    HMI_Message_Request : ARRAY[0..121] OF BOOL;  (* #HMI メッセージ表示要求; [0] 未使用; [1] 【Y616】A(左側) 供給スライド戻 異常表示; [2] 【Y617】A(左側) 供給スライド行 異常表示; [3] 【Y618】A(左側) 供給ピックアップ戻 異常表示; [4] 【Y619】A(左側) 供給ピックアップ行 異常表示; [5] 【Y620】A(左側) 供給チャック閉 戻 異常表示; [6] 【Y621】A(左側) 供給チャック開 行 異常表示; [7] 【Y622】B(右側) 供給スライド戻 異常表示; [8] 【Y623】B(右側) 供給スライド行 異常表示; [9] 【Y624】B(右側) 供給ピックアップ戻 異常表示; [10] 【Y625】B(右側) 供給ピックアップ行 異常表示; [11] 【Y626】B(右側) 供給チャック閉 戻 異常表示; [12] 【Y627】B(右側) 供給チャック開 行 異常表示; [13] 【Y700】A(左側) 高さ検査押え戻 異常表示; [14] 【Y701】A(左側) 高さ検査押え行 異常表示; [15] 【Y702】A(左側) 高さ検査持上戻 異常表示; [16] 【Y703】A(左側) 高さ検査持上行 異常表示; [17] 【Y704】A(左側) NG1ピックアップ戻 異常表示; [18] 【Y705】A(左側) NG1ピックアップ 行 異常表示; [19] 【Y706】A(左側) NG1チャック戻 異常表示; [20] 【Y707】A(左側) NG1チャック行 異常表示; [21] 【Y708】A(左側)ST4 反転1チャック閉 異常表示; [22] 【Y709】A(左側)ST4 反転1チャック開 異常表示; [23] 【Y710】A(左側)ST4 反転1ピックアップ戻 異常表示; [24] 【Y711】A(左側)ST4 反転1ピックアップ行 異常表示; [25] 【Y712】A(左側)ST6 反転2チャック閉 戻 異常表示; [26] 【Y713】A(左側)ST6 反転2チャック開 行 異常表示; [27] 【Y714】A(左側)ST6 反転2ピックアップ戻 異常表示; [28] 【Y715】A(左側)ST6 反転2ピックアップ行 異常表示; [29] 【Y716】A(左側) 排出チャック閉 戻 異常表示; [30] 【Y717】A(左側) 排出チャック開 行 異常表示; [31] 【Y718】A(左側) 排出フォルダ送り戻 異常表示; [32] 【Y719】A(左側) 排出フォルダ送り行 異常表示; [33] A(左側) 位置1ストッパー戻 異常表示; [34] 【Y720】A(左側) 位置1ストッパー 行 異常表示; [35] 【Y721】A(左側) 位置2ストッパー 異常表示; [36] 【Y721】A(左側) 位置2ストッパー 異常表示; [37] 【Y722】A(左側) 位置3ストッパー戻 異常表示; [38] 【Y722】A(左側) 位置3ストッパー行 異常表示; [39] Output_A_Error_M[33] 異常表示; [40] 【Y723】A(左側) 位置4ストッパー行 異常表示; [41] 【Y724】A(左側) 位置5ストッパー戻 異常表示; [42] 【Y724】A(左側) 位置5ストッパー行 異常表示; [43] 【Y725】A(左側) 位置6ストッパー戻 異常表示; [44] 【Y725】A(左側) 位置6ストッパー行 異常表示; [45] 【Y726】A(左側) ストックフォルダターン戻 異常表示; [46] 【Y727】A(左側) ストックフォルダターン行 異常表示; [47] 【Y728】A(左側) NG1仕分け 戻 異常表示; [48] 【Y729】A(左側) NG1仕分け 行 異常表示; [49] 【Y800】B(右側) 高さ検査押え戻 異常表示; [50] 【Y801】B(右側) 高さ検査押え行 異常表示; [51] 【Y802】B(右側) 高さ検査持上戻 異常表示; [52] 【Y803】B(右側) 高さ検査持上行 異常表示; [53] 【Y804】B(右側) NG1ピックアップ戻 異常表示; [54] 【Y805】B(右側) NG1ピックアップ 行 異常表示; [55] 【Y806】B(右側) NG1チャック戻 異常表示; [56] 【Y807】B(右側) NG1チャック行 異常表示; [57] 【Y808】B(右側)ST4 反転1チャック閉 戻 異常表示; [58] 【Y809】B(右側)ST4 反転1チャック開 戻 異常表示; [59] 【Y810】B(右側)ST4 反転1ピックアップ戻 異常表示; [60] 【Y811】B(右側)ST4 反転1ピックアップ行 異常表示; [61] 【Y812】B(右側)ST6 反転2チャック閉 戻 異常表示; [62] 【Y813】B(右側)ST6 反転2チャック開 行 異常表示; [63] 【Y814】B(右側)ST6 反転2ピックアップ戻 異常表示; [64] 【Y815】B(右側)ST6 反転2ピックアップ行 異常表示; [65] 【Y816】B(右側) 排出チャック閉 戻 異常表示; [66] 【Y817】B(右側) 排出チャック開 行 異常表示; [67] 【Y818】B(右側) 排出フォルダ送り戻 異常表示; [68] 【Y819】B(右側) 排出フォルダ送り行 異常表示; [69] 【Y820】B(右側) 位置1ストッパー 戻 異常表示; [70] 【Y820】B(右側) 位置1ストッパー 行 異常表示; [71] 【Y821】B(右側) 位置2ストッパー戻 異常表示; [72] 【Y821】B(右側) 位置2ストッパー行 異常表示; [73] 【Y822】B(右側) 位置3ストッパー戻 異常表示; [74] 【Y822】B(右側) 位置3ストッパー行 異常表示; [75] 【Y823】B(右側) 位置4ストッパー戻 異常表示; [76] 【Y823】B(右側) 位置4ストッパー行 異常表示; [77] 【Y824】B(右側) 位置5ストッパー戻 異常表示; [78] 【Y824】B(右側) 位置5ストッパー行 異常表示; [79] 【Y825】B(右側) 位置6ストッパー戻 異常表示; [80] 【Y825】B(右側) 位置6ストッパー行 異常表示; [81] 【Y826】B(右側) ストックフォルダターン戻 異常表示; [82] 【Y827】B(右側) ストックフォルダターン行 異常表示; [83] 【Y828】B(右側) NG1仕分け 戻 異常表示; [84] 【Y829】B(右側) NG1仕分け 行 異常表示; [85] 【Y1200】空コンテナ送り 戻 異常表示; [86] 【Y1201】空コンテナ送り 行 異常表示; [87] 【Y1202】段バラシ爪 戻 異常表示; [88] 【Y1203】段バラシ爪 行 異常表示; [89] 【Y1204】コンテナ排出 戻 異常表示; [90] 【Y1205】コンテナ排出 行 異常表示; [91] Output_Share_Error_M[7] 異常表示; [92] 【Y1207】箱入れチャック 行 異常表示; [93] 【Y1208】コンテナ仕分けストッパー 戻 異常表示; [94] 【Y1209】コンテナ仕分けストッパー 行 異常表示; [95] 【Y1210】コンテナ仕分け送り 戻 異常表示; [96] Output_Share_Error_M[12] 異常表示; [97] 【Y1300】A(左側) コンベア受渡送り戻 異常表示; [98] 【Y1301】A(左側) コンベア受渡送り行 異常表示; [99] 【Y1302】B(右側) コンベア受渡送り戻 異常表示; [100] 【Y1303】B(右側) コンベア受渡送り行 異常表示; [101] ST1 搬送ワーク不一致; [102] ST2 搬送ワーク不一致; [103] ST3 搬送ワーク不一致; [104] ST4 搬送ワーク不一致; [105] ST5 搬送ワーク不一致; [106] ST6 搬送ワーク不一致; [107] ST7 搬送ワーク不一致; [108] A(左側) ST1 FH測定時間超過; [109] A(左側) ST1 FH異常; [110] A(左側) ST5 FH異常; [111] B(右側) ST1 FH異常; [112] B(右側) ST5 FH異常; [113] A(左側) ST1 FH判定OK; [114] A(左側) ST1 FH判定NG1; [115] A(左側) ST1 FH判定NG2; [116] A(左側) ST1 検査前ワーク不一致; [117] A(左側) ST5 FH測定時間超過; [118] A(左側) ST5 FH判定OK; [119] A(左側) ST5 FH判定NG1; [120] A(左側) ST5 FH判定NG2; [121] A(左側) ST5 検査前ワーク不一致 *)
    HMI_Error_WorkSample : ARRAY[0..1] OF BOOL;  (* #HMI 再開前のワーク不一致; [0] A(左側) ST1; [1] A(左側) ST5 *)
    Error_ST1_A_Timeout : BOOL;  (* FHタイムアウト（非保持） *)
    Error_ST5_A_Timeout : BOOL;  (* FHタイムアウト（非保持） *)
    FH_B_ST1_Auto : BOOL;  (* B(右側) ST1 FH測定開始 *)
    Retry : ARRAY[0..99] OF BOOL;  (* 再試行：; [1] データ移動前 ワーク確; [4] ST3 検査前ワーク不一致エラー; [5] RCON1_1 機器異常; [6] A(左側) ST4 ワーク不一致エラー; [7] Stm A Axis000 絶対値位置決め エラー; [9] A(左側) ST6 ワーク不一致エラー; [10] Stm A Axis001 絶対値位置決め エラー; [12] RCON1_3 or 5機器異常 *)
    Stm_A_Rev_Axis000_MoveError : BOOL;  (* Stm A Axis000 絶対値位置決め エラー *)
    Stm_A_Rev1_Axis000_Power_Error : BOOL;  (* Stm A Axis000 サーボON エラー *)
    Stm_A_Rev_Axis001_MoveError : BOOL;  (* Stm A Axis001 絶対値位置決め エラー *)
    Stm_A_Rev2_Axis001_Power_Error : BOOL;  (* Stm A Axis001 サーボON エラー *)
    ST6_A_Rev2_End : BOOL;  (* ST6 A 動作完了 *)
    ST4_A_Rev_End : BOOL;  (* ST4 A 動作完了 *)
    RCON2_1_M : ARRAY[0..99] OF BOOL;  (* #RCON2_1 段バラシ; [1] 開始指令保持; [2] 予備 *)
    RCON2_1_IN_PositionDone : BOOL;  (* 位置決め完了 *)
    RCON2_1_IN_HomeDone : BOOL;  (* 原点復帰完了 *)
    RCON2_1_IN_Moving : BOOL;  (* 移動中 *)
    RCON2_1_IN_EmergencyStop : BOOL;  (* 非常停止状態（監視） *)
    RCON2_1_IN_ControllerReady : BOOL;  (* 準備完了 *)
    RCON2_1_IN_Zone2 : BOOL;  (* ゾーン2内 *)
    RCON2_1_IN_Zone1 : BOOL;  (* ゾーン1内 *)
    RCON2_1_IN_CommandDone : BOOL;  (* 指令完了 *)
    RCON2_1_IN_OverloadWarning : BOOL;  (* 過負荷警告 *)
    RCON2_1_IN_PushMiss : BOOL;  (* 押付け空振り（未使用） *)
    RCON2_1_IN_ServoReady : BOOL;  (* サーボON状態 *)
    RCON2_1_IN_Alarm : BOOL;  (* 軸異常 *)
    RCON2_1_Ready : BOOL;  (* 動作準備（安全許可とは別） *)
    RCON2_1_MoveDone : BOOL;  (* 動作完了 *)
    RCON2_1_OUT_TargetPos_mm : LREAL;  (* 目標位置 [mm] *)
    RCON2_1_OUT_PositionBand_mm : LREAL;  (* 位置決め幅 [mm] *)
    RCON2_1_OUT_Speed_mm_s : LREAL;  (* 指令速度 [mm/s] *)
    RCON2_1_OUT_AccDec_G : LREAL;  (* 加減速度 [G] *)
    RCON2_1_OUT_PushLimit_pct : LREAL;  (* 押付け制限 [%]（未使用） *)
    RCON2_1_ActualPos_mm : LREAL;  (* 現在位置 [mm] *)
    RCON2_1_Current_mA : DINT;  (* 指令電流 [mA]（監視値） *)
    RCON2_1_ActualSpeed_mm_s : LREAL;  (* 現在速度 [mm/s] *)
    RCON2_1_AlarmCode : UINT;  (* 軸異常コード *)
    RCON2_1_DataValid : BOOL;  (* 入力有効（安全許可とは別） *)
    RCON2_1_Auto : ARRAY[0..99] OF Bool;  (* 自動移動要求; [1] 初期動作① セイフティ; [2] 1段目 Pos; [3] 初期動作② セイフティ; [4] コンテナ排出 *)
    RCON2_2_M : ARRAY[0..99] OF BOOL;  (* #RCON2_2 箱詰めX; [1] 開始指令保持; [2] 今回移動受付：PEND OFF確認; [3] 自動開始許可 *)
    RCON2_2_IN_PositionDone : BOOL;  (* 位置決め完了 *)
    RCON2_2_IN_HomeDone : BOOL;  (* 原点復帰完了 *)
    RCON2_2_IN_Moving : BOOL;  (* 移動中 *)
    RCON2_2_IN_EmergencyStop : BOOL;  (* 非常停止状態（監視） *)
    RCON2_2_IN_ControllerReady : BOOL;  (* 準備完了 *)
    RCON2_2_IN_Zone2 : BOOL;  (* ゾーン2内 *)
    RCON2_2_IN_Zone1 : BOOL;  (* ゾーン1内 *)
    RCON2_2_IN_CommandDone : BOOL;  (* 指令完了 *)
    RCON2_2_IN_OverloadWarning : BOOL;  (* 過負荷警告 *)
    RCON2_2_IN_PushMiss : BOOL;  (* 押付け空振り（未使用） *)
    RCON2_2_IN_ServoReady : BOOL;  (* サーボON状態 *)
    RCON2_2_IN_Alarm : BOOL;  (* 軸異常 *)
    RCON2_2_Ready : BOOL;  (* 動作準備（安全許可とは別） *)
    RCON2_2_MoveDone : BOOL;  (* 動作完了 *)
    RCON2_2_OUT_TargetPos_mm : LREAL;  (* 目標位置 [mm] *)
    RCON2_2_OUT_PositionBand_mm : LREAL;  (* 位置決め幅 [mm] *)
    RCON2_2_OUT_Speed_mm_s : LREAL;  (* 指令速度 [mm/s] *)
    RCON2_2_OUT_AccDec_G : LREAL;  (* 加減速度 [G] *)
    RCON2_2_OUT_PushLimit_pct : LREAL;  (* 押付け制限 [%]（未使用） *)
    RCON2_2_ActualPos_mm : LREAL;  (* 現在位置 [mm] *)
    RCON2_2_Current_mA : DINT;  (* 指令電流 [mA]（監視値） *)
    RCON2_2_ActualSpeed_mm_s : LREAL;  (* 現在速度 [mm/s] *)
    RCON2_2_AlarmCode : UINT;  (* 軸異常コード *)
    RCON2_2_DataValid : BOOL;  (* 入力有効（安全許可とは別） *)
    RCON2_2_Auto : ARRAY[0..99] OF Bool;  (* 自動移動要求; [1] 自動要求1（未接続）; [2] 自動要求2（未接続）; [3] 自動要求3（未接続） *)
    RCON2_3_M : ARRAY[0..99] OF BOOL;  (* #RCON2_3 箱詰めY; [1] 開始指令保持; [2] 今回移動受付：PEND OFF確認; [3] 自動開始許可 *)
    RCON2_3_IN_PositionDone : BOOL;  (* 位置決め完了 *)
    RCON2_3_IN_HomeDone : BOOL;  (* 原点復帰完了 *)
    RCON2_3_IN_Moving : BOOL;  (* 移動中 *)
    RCON2_3_IN_EmergencyStop : BOOL;  (* 非常停止状態（監視） *)
    RCON2_3_IN_ControllerReady : BOOL;  (* 準備完了 *)
    RCON2_3_IN_Zone2 : BOOL;  (* ゾーン2内 *)
    RCON2_3_IN_Zone1 : BOOL;  (* ゾーン1内 *)
    RCON2_3_IN_CommandDone : BOOL;  (* 指令完了 *)
    RCON2_3_IN_OverloadWarning : BOOL;  (* 過負荷警告 *)
    RCON2_3_IN_PushMiss : BOOL;  (* 押付け空振り（未使用） *)
    RCON2_3_IN_ServoReady : BOOL;  (* サーボON状態 *)
    RCON2_3_IN_Alarm : BOOL;  (* 軸異常 *)
    RCON2_3_Ready : BOOL;  (* 動作準備（安全許可とは別） *)
    RCON2_3_MoveDone : BOOL;  (* 動作完了 *)
    RCON2_3_OUT_TargetPos_mm : LREAL;  (* 目標位置 [mm] *)
    RCON2_3_OUT_PositionBand_mm : LREAL;  (* 位置決め幅 [mm] *)
    RCON2_3_OUT_Speed_mm_s : LREAL;  (* 指令速度 [mm/s] *)
    RCON2_3_OUT_AccDec_G : LREAL;  (* 加減速度 [G] *)
    RCON2_3_OUT_PushLimit_pct : LREAL;  (* 押付け制限 [%]（未使用） *)
    RCON2_3_ActualPos_mm : LREAL;  (* 現在位置 [mm] *)
    RCON2_3_Current_mA : DINT;  (* 指令電流 [mA]（監視値） *)
    RCON2_3_ActualSpeed_mm_s : LREAL;  (* 現在速度 [mm/s] *)
    RCON2_3_AlarmCode : UINT;  (* 軸異常コード *)
    RCON2_3_DataValid : BOOL;  (* 入力有効（安全許可とは別） *)
    RCON2_3_Auto : ARRAY[0..99] OF Bool;  (* 自動移動要求; [1] 自動要求1（未接続）; [2] 自動要求2（未接続）; [3] 自動要求3（未接続） *)
    RCON2_4_M : ARRAY[0..99] OF BOOL;  (* #RCON2_4 箱詰めZ; [1] 開始指令保持; [2] 今回移動受付：PEND OFF確認; [3] 自動開始許可 *)
    RCON2_4_IN_PositionDone : BOOL;  (* 位置決め完了 *)
    RCON2_4_IN_HomeDone : BOOL;  (* 原点復帰完了 *)
    RCON2_4_IN_Moving : BOOL;  (* 移動中 *)
    RCON2_4_IN_EmergencyStop : BOOL;  (* 非常停止状態（監視） *)
    RCON2_4_IN_ControllerReady : BOOL;  (* 準備完了 *)
    RCON2_4_IN_Zone2 : BOOL;  (* ゾーン2内 *)
    RCON2_4_IN_Zone1 : BOOL;  (* ゾーン1内 *)
    RCON2_4_IN_CommandDone : BOOL;  (* 指令完了 *)
    RCON2_4_IN_OverloadWarning : BOOL;  (* 過負荷警告 *)
    RCON2_4_IN_PushMiss : BOOL;  (* 押付け空振り（未使用） *)
    RCON2_4_IN_ServoReady : BOOL;  (* サーボON状態 *)
    RCON2_4_IN_Alarm : BOOL;  (* 軸異常 *)
    RCON2_4_Ready : BOOL;  (* 動作準備（安全許可とは別） *)
    RCON2_4_MoveDone : BOOL;  (* 動作完了 *)
    RCON2_4_OUT_TargetPos_mm : LREAL;  (* 目標位置 [mm] *)
    RCON2_4_OUT_PositionBand_mm : LREAL;  (* 位置決め幅 [mm] *)
    RCON2_4_OUT_Speed_mm_s : LREAL;  (* 指令速度 [mm/s] *)
    RCON2_4_OUT_AccDec_G : LREAL;  (* 加減速度 [G] *)
    RCON2_4_OUT_PushLimit_pct : LREAL;  (* 押付け制限 [%]（未使用） *)
    RCON2_4_ActualPos_mm : LREAL;  (* 現在位置 [mm] *)
    RCON2_4_Current_mA : DINT;  (* 指令電流 [mA]（監視値） *)
    RCON2_4_ActualSpeed_mm_s : LREAL;  (* 現在速度 [mm/s] *)
    RCON2_4_AlarmCode : UINT;  (* 軸異常コード *)
    RCON2_4_DataValid : BOOL;  (* 入力有効（安全許可とは別） *)
    RCON2_4_Auto : ARRAY[0..99] OF Bool;  (* 自動移動要求; [1] 自動要求1（未接続）; [2] 自動要求2（未接続）; [3] 自動要求3（未接続） *)
    RCON2_5_M : ARRAY[0..99] OF BOOL;  (* #RCON2_5 コンテナ設置; [1] 開始指令保持; [2] 今回移動受付：PEND OFF確認; [3] 自動開始許可 *)
    RCON2_5_IN_PositionDone : BOOL;  (* 位置決め完了 *)
    RCON2_5_IN_HomeDone : BOOL;  (* 原点復帰完了 *)
    RCON2_5_IN_Moving : BOOL;  (* 移動中 *)
    RCON2_5_IN_EmergencyStop : BOOL;  (* 非常停止状態（監視） *)
    RCON2_5_IN_ControllerReady : BOOL;  (* 準備完了 *)
    RCON2_5_IN_Zone2 : BOOL;  (* ゾーン2内 *)
    RCON2_5_IN_Zone1 : BOOL;  (* ゾーン1内 *)
    RCON2_5_IN_CommandDone : BOOL;  (* 指令完了 *)
    RCON2_5_IN_OverloadWarning : BOOL;  (* 過負荷警告 *)
    RCON2_5_IN_PushMiss : BOOL;  (* 押付け空振り（未使用） *)
    RCON2_5_IN_ServoReady : BOOL;  (* サーボON状態 *)
    RCON2_5_IN_Alarm : BOOL;  (* 軸異常 *)
    RCON2_5_Ready : BOOL;  (* 動作準備（安全許可とは別） *)
    RCON2_5_MoveDone : BOOL;  (* 動作完了 *)
    RCON2_5_OUT_TargetPos_mm : LREAL;  (* 目標位置 [mm] *)
    RCON2_5_OUT_PositionBand_mm : LREAL;  (* 位置決め幅 [mm] *)
    RCON2_5_OUT_Speed_mm_s : LREAL;  (* 指令速度 [mm/s] *)
    RCON2_5_OUT_AccDec_G : LREAL;  (* 加減速度 [G] *)
    RCON2_5_OUT_PushLimit_pct : LREAL;  (* 押付け制限 [%]（未使用） *)
    RCON2_5_ActualPos_mm : LREAL;  (* 現在位置 [mm] *)
    RCON2_5_Current_mA : DINT;  (* 指令電流 [mA]（監視値） *)
    RCON2_5_ActualSpeed_mm_s : LREAL;  (* 現在速度 [mm/s] *)
    RCON2_5_AlarmCode : UINT;  (* 軸異常コード *)
    RCON2_5_DataValid : BOOL;  (* 入力有効（安全許可とは別） *)
    RCON2_5_Auto : ARRAY[0..99] OF Bool;  (* 自動移動要求; [1] コンテナトレイ方向NG; [2] 自動要求2（未接続）; [3] 自動要求3（未接続） *)
    Auto_Com_Start : BOOL;  (* 共通ユニット自動運転開始 *)
    Destacker_M : ARRAY[0..99] OF Bool;  (* 段バラシ工程; [5] 初回安全位置なし; [4] 初回安全位置あり; [2] 初回の爪保持; [3] 初回の位置判定; [6] 初回の爪戻し; [26] 初回確認済み; [27] 初回安全 前完了解除; [28] 初回1段 前完了解除; [29] 初回戻り 前完了解除; [30] 1段目 前完了解除; [31] 2段目 前完了解除; [32] 排出 前完了解除; [1] 初回確認開始; [7] 初回安全位置移動; [8] 初回1段目移動; [9] 初回コンテナ保持; [10] 初回安全位置戻り; [11] 初回の送り戻し; [12] 通常サイクル開始; [13] 送り戻り待ち; [14] コンテナ確認中; [15] コンテナ確認OK; [16] 1段目位置へ移動; [17] コンテナ切り離し; [18] 段積み判定; [19] 2段以上; [20] 1段のみ; [21] 2段目位置へ移動; [22] 上段コンテナ保持; [23] 安全・排出位置移動; [24] 送り行待ち; [25] 送り戻り待ち *)
    HMI_RCON2_1_OUT_TargetPos : ARRAY[0..99] OF LREAL;  (* 段バラシ 目標位置 [mm]; [1] ①④セイフティ・排出 Pos; [2] ②1段目 Pos; [3] ③2段目 Pos *)
    BoxPacking_Busy : BOOL;  (* 箱詰め動作中 *)
    Destacker_End : BOOL;  (* 1サイクル完了 *)
    Destacker_Error : BOOL;  (* 方向・1段目確認異常 *)
    Error_Destacker_M : ARRAY[0..99] OF Bool;  (* 段バラシエラー： *)
    ST7_B_SF_Wait_Pickup : BOOL;  (* フォルダストックB取出し待ち *)
END_VAR
VAR_GLOBAL RETAIN
    HMI_A_SF_StackPitch_mm : LREAL;  (* 左SF積みピッチ [mm] *)
END_VAR
VAR_GLOBAL
    A_Total_CT : INT;  (* A(左側)生産数 *)
    HMI_RCON2_4_OUT_TargetPos : ARRAY[0..99] OF LREAL;  (* 箱詰めZ：; [1] セイフティ 上昇 Pos; [2] フォルダストック 取出し降下Pos; [3] トレイ ワーク梱包 降下Pos *)
    Box_Total_CT : INT;  (* コンテナ入数 *)
END_VAR
VAR_GLOBAL RETAIN
    HMI_Box_X_Pitch_mm : LREAL;  (* 箱詰めX方向の1ピッチ [mm]：符号付き。正=座標増、負=座標減。使用前に設定。 *)
    HMI_Box_Y_Pitch_mm : LREAL;  (* 箱詰めY方向の1ピッチ [mm]：符号付き。正=座標増、負=座標減。使用前に設定。 *)
END_VAR

PROGRAM ModeManagement_モード管理
VAR
    Setting_M : BOOL;
    Manual_M : BOOL;
    Auto_M : BOOL;
    Dummy_M : BOOL;
    Inital_M : BOOL;
    Output_Error_M : ARRAY[0..99] OF Bool;
    Index_Error_001 : DINT;
    Index_B_001 : DINT;
    Index_Share_001 : DINT;
    Error_TON : ARRAY[0..99] OF TON;  (* [2] A(左側) ST1 測定タイムアウト; [4] A(左側) ST5 測定タイムアウト *)
    Error_TOF : ARRAY[0..99] OF TOF;
    AutoMode_A_M : ARRAY[0..99] OF Bool;
    ６ : DINT;
    ST4_A_Rev_01_Origin_M : ARRAY[0..99] OF Bool;  (* A(左側) ST4 反転1 原点復帰工程; [1] A(左側) ST4 反転1 原点復帰開始; [2] A(左側) ST4 反転1 原点復帰中; [3] A(左側) ST4 反転1 ピックアップ戻; [4] A(左側) ST4 反転1 モータ原点復帰開始; [5] A(左側) ST4 反転1 ピックアップ行; [6] A(左側) ST4 反転1 チャック閉; [7] A(左側) ST4 反転1 原点復帰完了（ワーク無） *)
    ST4_A_Rev_01_OriginDone : BOOL;  (* A(左側) ST4 反転1 原点復帰完了 *)
    ST4_A_Rev_02_Origin_M : ARRAY[0..99] OF Bool;  (* A(左側) ST6 反転2 原点復帰工程; [1] A(左側) ST6 反転2 原点復帰開始; [2] A(左側) ST6 反転2 原点復帰中; [3] A(左側) ST6 反転2 ピックアップ戻; [4] A(左側) ST6 反転2 モータ原点復帰開始; [5] A(左側) ST6 反転2 ピックアップ行; [6] A(左側) ST6 反転2 チャック閉; [7] A(左側) ST6 反転2 原点復帰完了（ワーク無） *)
    ST4_A_Rev_02_OriginDone : BOOL;  (* A(左側) ST6 反転2 原点復帰完了 *)
    ST4_B_Rev_01_Origin_M : ARRAY[0..99] OF Bool;  (* B(右側) ST4 反転1 原点復帰工程; [1] B(右側) ST4 反転1 原点復帰開始; [2] B(右側) ST4 反転1 原点復帰中; [3] B(右側) ST4 反転1 ピックアップ戻; [4] B(右側) ST4 反転1 モータ原点復帰開始; [5] B(右側) ST4 反転1 ピックアップ行; [6] B(右側) ST4 反転1 チャック閉; [7] B(右側) ST4 反転1 原点復帰完了（ワーク無） *)
    ST4_B_Rev_01_OriginDone : BOOL;  (* B(右側) ST4 反転1 原点復帰完了 *)
    ST4_B_Rev_02_Origin_M : ARRAY[0..99] OF Bool;  (* B(右側) ST6 反転2 原点復帰工程; [1] B(右側) ST6 反転2 原点復帰開始; [2] B(右側) ST6 反転2 原点復帰中; [3] B(右側) ST6 反転2 ピックアップ戻; [4] B(右側) ST6 反転2 モータ原点復帰開始; [5] B(右側) ST6 反転2 ピックアップ行; [6] B(右側) ST6 反転2 チャック閉; [7] B(右側) ST6 反転2 原点復帰完了（ワーク無） *)
    ST4_B_Rev_02_OriginDone : BOOL;  (* B(右側) ST6 反転2 原点復帰完了 *)
    ST1_B_Ca1_M : BOOL;
END_VAR
VAR_EXTERNAL
    Output_A_Error_M : ARRAY[0..99] OF Bool;
    Output_A_Restart_M : ARRAY[0..99] OF Bool;
    In_Sw_RESET : BOOL;
    In_Sw_START : BOOL;
    ManualMode : BOOL;
    M9999 : BOOL;
    Output_B_Error_M : ARRAY[0..99] OF Bool;  (* B(右側)シリンダエラー *)
    Output_B_Restart_M : ARRAY[0..99] OF Bool;  (* B(右側)シリンダ再開： *)
    Output_Share_Error_M : ARRAY[0..99] OF Bool;
    Output_Share_Restart_M : ARRAY[0..99] OF Bool;
    TimerQ_In_Sen_Accum_CV_A_Full : BOOL;
    Out_TDC_Stop : BOOL;
    In_Sen_Unl_Conv_A_Pass : BOOL;
    In_Sen_Accum_CV_A_Full : BOOL;
    In_Sen_Unl_Conv_B_Pass : BOOL;
    Pause : ARRAY[0..99] OF Bool;  (* [3] FH A(左側) ST1; [9] FH A(左側) ST5; [10] FH B(右側) ST1; [11] FH B(右側) ST5; [12] A(左側) ST6 反転2 ワーク不一致 *)
    AutoMode : BOOL;
    In_Sen_DOOR_01 : BOOL;
    In_Sen_DOOR_02 : BOOL;
    In_Sen_DOOR_03 : BOOL;
    In_Sen_DOOR_04 : BOOL;
    In_Sen_DOOR_05 : BOOL;
    In_Sen_DOOR_06 : BOOL;
    In_Sw_EMS1 : BOOL;
    In_Sw_EMS2 : BOOL;
    In_Sw_EMS3 : BOOL;
    In_Sen_AIR１_Pressure_01 : BOOL;
    In_Sen_AIR１_Pressure_02 : BOOL;
    In_Sen_AIR１_Pressure_03 : BOOL;
    TEST_M : ARRAY[0..99] OF Bool;
    ST0_Sup_Start : BOOL;  (* ST0_動作開始 *)
    Out_CYw_Sply_Pick_A_H_Auto : ARRAY[0..10] OF Bool;
    Out_CYw_Sply_Pick_A_H_Done : BOOL;
    Out_CYw_Sply_Slide_A_H_Auto : ARRAY[0..10] OF Bool;
    Out_CYw_Sply_Slide_A_H_Done : BOOL;
    Out_CYw_Sup_Chuck_A_Cl_H_Auto : ARRAY[0..10] OF Bool;
    Out_CYw_Sup_Chuck_A_Cl_H_Done : BOOL;
    In_Sen_Accum_CV_A_Arrival : BOOL;
    In_Sen_Work_A_Pos_00 : BOOL;
    Out_CYw_Sply_Pick_A_F_Auto : ARRAY[0..10] OF Bool;
    Out_CYw_Sply_Pick_A_F_Done : BOOL;
    Out_CYw_Sup_Chuck_A_Cl_F_Auto : ARRAY[0..10] OF Bool;
    Out_CYw_Sup_Chuck_A_Cl_F_Done : BOOL;
    Out_CYw_Sply_Slide_A_F_Auto : ARRAY[0..10] OF Bool;
    Out_CYw_Sply_Slide_A_F_Done : BOOL;
    Ins_A_Cv_Error : BOOL;
    Station_A_Data : ARRAY[0..8] OF sData;
    Ins_A_Cv_M : ARRAY[0..99] OF Bool;
    HMI_MessageNo : ARRAY[0..9] OF UINT;
    FH_A_ST1_Auto : BOOL;
    In_Sen_Accum_CV_B_Full : BOOL;
    FH_Line3_Error_Status_1 : BOOL;
    FH_Line0_Error_Status_1 : BOOL;
    FH_Line1_Error_Status_1 : BOOL;
    FH_Line2_Error_Status_1 : BOOL;
    FH_Line0_Error_Clear_1 : BOOL;
    FH_Line1_Error_Clear_1 : BOOL;
    FH_Line2_Error_Clear_1 : BOOL;
    FH_Line3_Error_Clear_1 : BOOL;
    Ins_A_Next_Cycle : BOOL;
    OriginDone : BOOL;  (* 原点復帰完了 *)
    DummyDone : BOOL;  (* ダミーチェック完了 *)
    HMI_CurrentPage : STRING[256];
    Ins_A_End : BOOL;
    Auto_A_Start : BOOL;  (* 自動運転 開始 *)
    Auto_Ready : BOOL;  (* 自動運転可能 *)
    ST0_A_Sup_Busy : BOOL;
    ST1_A_Ca1_Busy : BOOL;
    RCON1_1_IN_Alarm : BOOL;  (* 軸異常 *)
    RCON1_1_IN_EmergencyStop : BOOL;  (* 非常停止状態（監視） *)
    RCON1_1_Error : BOOL;  (* 異常予備（未接続） *)
    RCON1_1_IN_HomeDone : BOOL;  (* 原点復帰完了 *)
    RCON1_1_Error_Clear : BOOL;  (* 解除予備（未接続） *)
    Error_M : ARRAY[0..99] OF Bool;  (* エラー：; [1] シリンダ; [2] コンベア＆ドアセンサ; [3] 未使用：Error_ST1_A_M[0]へ移行; [4] A(左側)検査コンベア ワーク不一致; [5] 未使用：Error_ST3_A_M[1]へ移行; [9] 未使用：Error_ST5_A_M[0]へ移行; [10] 未使用：Error_ST1_B_M[0]へ移行; [11] 未使用：Error_ST5_B_M[0]へ移行; [12] 未使用：Error_ST6_A_M[0]へ移行 *)
    ST1_A_Ca1_M : ARRAY[0..99] OF Bool;  (* [6] A(左側) ST1 検査前ワーク不一致 *)
    ST2_A_Hgt_M : ARRAY[0..99] OF Bool;
    ST3_A_Dis1_M : ARRAY[0..99] OF Bool;
    HMI_Home_SW : BOOL;
    Origin_Busy : BOOL;  (* 原点復帰中 *)
    Out_CYw_Rev_01_Pick_A_H_Origin : ARRAY[0..10] OF Bool;  (* 原点復帰【Y710】A(左側)ST4 反転1ピックアップ戻： *)
    Out_CYw_Rev_01_Pick_A_H_Done : BOOL;  (* 【Y710】A(左側)ST4 反転1ピックアップ戻 動作完了 *)
    Stm_A_Rev_Axis000_Origin : BOOL;  (* A(左側) ST4 反転1 モータ原点復帰開始 *)
    Stm_A_Rev_Axis000_OriginDone : BOOL;  (* A(左側) ST4 反転1 モータ原点復帰完了 *)
    Out_CYw_Rev_01_Pick_A_F_Origin : ARRAY[0..99] OF Bool;  (* 原点復帰【Y711】A(左側)ST4 反転1ピックアップ行： *)
    Out_CYw_Rev_01_Pick_A_F_Done : BOOL;  (* 【Y711】A(左側)ST4 反転1ピックアップ行 動作完了 *)
    Out_CYw_Rev_01_Chk_A_H_Origin : ARRAY[0..99] OF Bool;  (* 原点復帰【Y708】A(左側)ST4 反転1チャック閉： *)
    Out_CYw_Rev_01_Chk_A_H_Done : BOOL;  (* 【Y708】A(左側)ST4 反転1チャック閉 動作完了 *)
    TimerQ_In_Sen_Work_A_Pos_04 : BOOL;
    Out_CYw_Rev_02_Pick_A_H_Origin : ARRAY[0..10] OF Bool;  (* 原点復帰 【Y714】A(左側)ST6 反転2ピックアップ戻 *)
    Out_CYw_Rev_02_Pick_A_H_Done : BOOL;  (* 【Y714】A(左側)ST6 反転2ピックアップ戻 動作完了 *)
    Stm_A_Rev_Axis001_Origin : BOOL;  (* A(左側) ST6 反転2 モータ原点復帰開始 *)
    Stm_A_Rev_Axis001_OriginDone : BOOL;  (* A(左側) ST6 反転2 モータ原点復帰完了 *)
    Out_CYw_Rev_02_Pick_A_F_Origin : ARRAY[0..99] OF Bool;  (* 原点復帰 【Y715】A(左側)ST6 反転2ピックアップ行 *)
    Out_CYw_Rev_02_Pick_A_F_Done : BOOL;  (* 【Y715】A(左側)ST6 反転2ピックアップ行 動作完了 *)
    Out_CYw_Rev_02_Chk_A_H_Origin : ARRAY[0..99] OF Bool;  (* 原点復帰 【Y712】A(左側)ST6 反転2チャック閉 戻 *)
    Out_CYw_Rev_02_Chk_A_H_Done : BOOL;  (* 【Y712】A(左側)ST6 反転2チャック閉 戻 動作完了 *)
    TimerQ_In_Sen_Work_A_Pos_06 : BOOL;  (* 【X208】A(左側)ワーク位置6 *)
    Auto_B_Start : BOOL;  (* B(右側)自動運転開始（後続処理未接続） *)
    Out_CYw_Rev_01_Pick_B_H_Origin : ARRAY[0..10] OF Bool;  (* 原点復帰 【Y810】B(右側)ST4 反転1ピックアップ戻 *)
    Out_CYw_Rev_01_Pick_B_H_Done : BOOL;  (* 【Y810】B(右側)ST4 反転1ピックアップ戻 動作完了 *)
    Stm_B_Rev_Axis002_Origin : BOOL;  (* B(右側) ST4 反転1 モータ原点復帰開始 *)
    Stm_B_Rev_Axis002_OriginDone : BOOL;  (* B(右側) ST4 反転1 モータ原点復帰完了 *)
    Out_CYw_Rev_01_Pick_B_F_Origin : ARRAY[0..99] OF Bool;  (* 原点復帰 【Y811】B(右側)ST4 反転1ピックアップ行 *)
    Out_CYw_Rev_01_Pick_B_F_Done : BOOL;  (* 【Y811】B(右側)ST4 反転1ピックアップ行 動作完了 *)
    Out_CYw_Rev_01_Chk_B_H_Origin : ARRAY[0..99] OF Bool;  (* 原点復帰 【Y808】B(右側)ST4 反転1チャック閉 戻 *)
    Out_CYw_Rev_01_Chk_B_H_Done : BOOL;  (* 【Y808】B(右側)ST4 反転1チャック閉 戻 動作完了 *)
    TimerQ_In_Sen_Work_B_Pos_04 : BOOL;  (* 【X406】B(右側)ワーク位置4 *)
    Out_CYw_Rev_02_Pick_B_H_Origin : ARRAY[0..10] OF Bool;  (* 原点復帰 【Y814】B(右側)ST6 反転2ピックアップ戻 *)
    Out_CYw_Rev_02_Pick_B_H_Done : BOOL;  (* 【Y814】B(右側)ST6 反転2ピックアップ戻 動作完了 *)
    Stm_B_Rev_Axis003_Origin : BOOL;  (* B(右側) ST6 反転2 モータ原点復帰開始 *)
    Stm_B_Rev_Axis003_OriginDone : BOOL;  (* B(右側) ST6 反転2 モータ原点復帰完了 *)
    Out_CYw_Rev_02_Pick_B_F_Origin : ARRAY[0..99] OF Bool;  (* 原点復帰 【Y815】B(右側)ST6 反転2ピックアップ行 *)
    Out_CYw_Rev_02_Pick_B_F_Done : BOOL;  (* 【Y815】B(右側)ST6 反転2ピックアップ行 動作完了 *)
    Out_CYw_Rev_02_Chk_B_H_Origin : ARRAY[0..99] OF Bool;  (* 原点復帰 【Y812】B(右側)ST6 反転2チャック閉 戻 *)
    Out_CYw_Rev_02_Chk_B_H_Done : BOOL;  (* 【Y812】B(右側)ST6 反転2チャック閉 戻 動作完了 *)
    TimerQ_In_Sen_Work_B_Pos_06 : BOOL;  (* 【X408】B(右側)ワーク位置6 *)
    ST4_A_Rev1_M : ARRAY[0..99] OF Bool;  (* [10] A(左側) ST4 ワーク不一致エラー; [12] 【Y708】A(左側) ST4 反転1チャック閉 *)
    ST5_A_Ca2_M : ARRAY[0..99] OF Bool;  (* A(左側) ST5 カメラ2工程; [1] A(左側) ST5 カメラ2検査開始; [2] 【Y724】A(左側) ST5 ストッパー戻; [3] A(左側) ST5 ワーク有無判定; [4] A(左側) ST5 ワーク有; [5] A(左側) ST5 ワーク無; [6] A(左側) ST5 検査前ワーク不一致; [7] A(左側) ST5 FH測定開始 *)
    FH_A_ST5_Auto : BOOL;  (* A(左側) ST5 FH自動測定 *)
END_VAR
VAR_EXTERNAL CONSTANT
    ST6_A_Rev2_M : ARRAY[0..99] OF Bool;  (* A(左側) ST6 反転2工程; [1] A(左側) ST6 反転2 動作開始; [2] A(左側) ST6 反転2 【Y714】ピックアップ戻; [3] A(左側) ST6 反転2 【Y725】位置6ストッパー戻; [4] A(左側) ST6 反転2 原点角度転送; [5] A(左側) ST6 反転2 原点位置移動開始; [6] A(左側) ST6 反転2 原点位置移動完了; [7] A(左側) ST6 反転2 ワーク有無判定; [8] A(左側) ST6 反転2 ワーク有・前工程OK; [9] A(左側) ST6 反転2 ワーク無・前工程NG; [10] A(左側) ST6 反転2 ワーク不一致エラー; [11] A(左側) ST6 反転2 【Y715】反転前ピックアップ行; [12] A(左側) ST6 反転2 【Y712】チャック閉; [13] A(左側) ST6 反転2 【Y714】反転前ピックアップ戻; [14] A(左側) ST6 反転2 反転角度転送; [15] A(左側) ST6 反転2 反転位置移動完了; [16] A(左側) ST6 反転2 【Y715】設置ピックアップ行; [17] A(左側) ST6 反転2 【Y713】チャック開; [18] A(左側) ST6 反転2 【Y714】設置ピックアップ戻 *)
END_VAR
VAR_EXTERNAL
    ST7_A_Dis2_M : ARRAY[0..99] OF Bool;  (* [9] ワーク有; [10] ワーク無; [11] 有無・NG満杯異常; [12] 回収下降位置転送; [13] 回収下降要求; [14] ワーク保持; [15] 保持後上昇位置転送; [16] 保持後上昇要求; [17] 仕分け位置選択; [18] OK選択; [19] キズNG選択; [20] 姿NG選択; [21] OK送り行開始; [22] 仕分け左右移動中; [23] 下降位置選択; [24] OK積み位置; [25] キズNG下降位置; [26] 姿NG下降位置; [27] 配置下降要求; [28] ワーク解放; [29] 解放後上昇位置転送; [30] 解放後上昇要求; [31] 左右原点位置転送; [32] 左右原点移動要求; [33] 最後の送り戻; [1] 排出動作開始; [2] 初期チャック戻; [3] 初期上昇位置転送; [4] 初期上昇要求; [5] 初期左右位置転送; [6] 初期左右移動要求; [7] 初期送り戻; [8] ワーク有無判定; [42] 今回ワーク加算済み; [43] 積み設定・判定異常; [44] フォルダ回転異常; [45] ワーク回収開始許可; [46] 今回の初期位置確認済み; [34] 初期上昇 前完了解除; [35] 初期左右 前完了解除; [36] 回収下降 前完了解除; [37] 保持後上昇 前完了解除; [38] 仕分け左右 前完了解除; [39] 配置下降 前完了解除; [40] 解放後上昇 前完了解除; [41] 左右戻り 前完了解除 *)
    Error_ST1_A_M : ARRAY[0..4] OF BOOL;  (* #A(左側) ST1 カメラ1 異常; [0] 総合異常; [1] 機器異常; [2] タイムアウト; [3] ワーク不一致; [4] 予備（監視なし） *)
    Error_ST1_B_M : ARRAY[0..4] OF BOOL;  (* #B(右側) ST1 カメラ1 異常; [0] 総合異常; [1] 機器異常; [2] 予備（監視なし）; [3] 予備（監視なし）; [4] 予備（監視なし） *)
    Error_ST2_A_M : ARRAY[0..4] OF BOOL;  (* #A(左側) ST2 高さ検査 異常; [0] 総合異常; [1] 予備（監視なし）; [2] 予備（監視なし）; [3] ワーク不一致; [4] 予備（監視なし） *)
    Error_ST3_A_M : ARRAY[0..4] OF BOOL;  (* #A(左側) ST3 NG1排出 異常; [0] 総合異常; [1] 機器異常; [2] 予備（監視なし）; [3] ワーク不一致; [4] 予備（監視なし） *)
    Error_ST4_A_M : ARRAY[0..4] OF BOOL;  (* #A(左側) ST4 反転1 異常; [0] 総合異常; [1] 予備（監視なし）; [2] 予備（監視なし）; [3] ワーク不一致; [4] 予備（監視なし） *)
    Error_ST5_A_M : ARRAY[0..4] OF BOOL;  (* #A(左側) ST5 カメラ2 異常; [0] 総合異常; [1] 機器異常; [2] タイムアウト; [3] ワーク不一致; [4] 予備（監視なし） *)
    Error_ST5_B_M : ARRAY[0..4] OF BOOL;  (* #B(右側) ST5 カメラ2 異常; [0] 総合異常; [1] 機器異常; [2] 予備（監視なし）; [3] 予備（監視なし）; [4] 予備（監視なし） *)
    Error_ST6_A_M : ARRAY[0..4] OF BOOL;  (* #A(左側) ST6 反転2 異常; [0] 総合異常; [1] 予備（監視なし）; [2] 予備（監視なし）; [3] ワーク不一致; [4] 予備（監視なし） *)
    Error_ST7_A_M : ARRAY[0..4] OF BOOL;  (* #A(左側) ST7 SF排出 異常; [0] 総合異常; [1] 予備（監視なし）; [2] 予備（監視なし）; [3] ワーク不一致; [4] 満杯 *)
    Error_ST7_A_Source_M : ARRAY[0..4] OF BOOL;  (* #A(左側) ST7 発生理由（内部保持）; [3] ワーク不一致; [4] 満杯（既存B側入力） *)
    HMI_Message_Request : ARRAY[0..121] OF BOOL;  (* #HMI メッセージ表示要求; [0] 未使用; [1] 【Y616】A(左側) 供給スライド戻 異常表示; [2] 【Y617】A(左側) 供給スライド行 異常表示; [3] 【Y618】A(左側) 供給ピックアップ戻 異常表示; [4] 【Y619】A(左側) 供給ピックアップ行 異常表示; [5] 【Y620】A(左側) 供給チャック閉 戻 異常表示; [6] 【Y621】A(左側) 供給チャック開 行 異常表示; [7] 【Y622】B(右側) 供給スライド戻 異常表示; [8] 【Y623】B(右側) 供給スライド行 異常表示; [9] 【Y624】B(右側) 供給ピックアップ戻 異常表示; [10] 【Y625】B(右側) 供給ピックアップ行 異常表示; [11] 【Y626】B(右側) 供給チャック閉 戻 異常表示; [12] 【Y627】B(右側) 供給チャック開 行 異常表示; [13] 【Y700】A(左側) 高さ検査押え戻 異常表示; [14] 【Y701】A(左側) 高さ検査押え行 異常表示; [15] 【Y702】A(左側) 高さ検査持上戻 異常表示; [16] 【Y703】A(左側) 高さ検査持上行 異常表示; [17] 【Y704】A(左側) NG1ピックアップ戻 異常表示; [18] 【Y705】A(左側) NG1ピックアップ 行 異常表示; [19] 【Y706】A(左側) NG1チャック戻 異常表示; [20] 【Y707】A(左側) NG1チャック行 異常表示; [21] 【Y708】A(左側)ST4 反転1チャック閉 異常表示; [22] 【Y709】A(左側)ST4 反転1チャック開 異常表示; [23] 【Y710】A(左側)ST4 反転1ピックアップ戻 異常表示; [24] 【Y711】A(左側)ST4 反転1ピックアップ行 異常表示; [25] 【Y712】A(左側)ST6 反転2チャック閉 戻 異常表示; [26] 【Y713】A(左側)ST6 反転2チャック開 行 異常表示; [27] 【Y714】A(左側)ST6 反転2ピックアップ戻 異常表示; [28] 【Y715】A(左側)ST6 反転2ピックアップ行 異常表示; [29] 【Y716】A(左側) 排出チャック閉 戻 異常表示; [30] 【Y717】A(左側) 排出チャック開 行 異常表示; [31] 【Y718】A(左側) 排出フォルダ送り戻 異常表示; [32] 【Y719】A(左側) 排出フォルダ送り行 異常表示; [33] A(左側) 位置1ストッパー戻 異常表示; [34] 【Y720】A(左側) 位置1ストッパー 行 異常表示; [35] 【Y721】A(左側) 位置2ストッパー 異常表示; [36] 【Y721】A(左側) 位置2ストッパー 異常表示; [37] 【Y722】A(左側) 位置3ストッパー戻 異常表示; [38] 【Y722】A(左側) 位置3ストッパー行 異常表示; [39] Output_A_Error_M[33] 異常表示; [40] 【Y723】A(左側) 位置4ストッパー行 異常表示; [41] 【Y724】A(左側) 位置5ストッパー戻 異常表示; [42] 【Y724】A(左側) 位置5ストッパー行 異常表示; [43] 【Y725】A(左側) 位置6ストッパー戻 異常表示; [44] 【Y725】A(左側) 位置6ストッパー行 異常表示; [45] 【Y726】A(左側) ストックフォルダターン戻 異常表示; [46] 【Y727】A(左側) ストックフォルダターン行 異常表示; [47] 【Y728】A(左側) NG1仕分け 戻 異常表示; [48] 【Y729】A(左側) NG1仕分け 行 異常表示; [49] 【Y800】B(右側) 高さ検査押え戻 異常表示; [50] 【Y801】B(右側) 高さ検査押え行 異常表示; [51] 【Y802】B(右側) 高さ検査持上戻 異常表示; [52] 【Y803】B(右側) 高さ検査持上行 異常表示; [53] 【Y804】B(右側) NG1ピックアップ戻 異常表示; [54] 【Y805】B(右側) NG1ピックアップ 行 異常表示; [55] 【Y806】B(右側) NG1チャック戻 異常表示; [56] 【Y807】B(右側) NG1チャック行 異常表示; [57] 【Y808】B(右側)ST4 反転1チャック閉 戻 異常表示; [58] 【Y809】B(右側)ST4 反転1チャック開 戻 異常表示; [59] 【Y810】B(右側)ST4 反転1ピックアップ戻 異常表示; [60] 【Y811】B(右側)ST4 反転1ピックアップ行 異常表示; [61] 【Y812】B(右側)ST6 反転2チャック閉 戻 異常表示; [62] 【Y813】B(右側)ST6 反転2チャック開 行 異常表示; [63] 【Y814】B(右側)ST6 反転2ピックアップ戻 異常表示; [64] 【Y815】B(右側)ST6 反転2ピックアップ行 異常表示; [65] 【Y816】B(右側) 排出チャック閉 戻 異常表示; [66] 【Y817】B(右側) 排出チャック開 行 異常表示; [67] 【Y818】B(右側) 排出フォルダ送り戻 異常表示; [68] 【Y819】B(右側) 排出フォルダ送り行 異常表示; [69] 【Y820】B(右側) 位置1ストッパー 戻 異常表示; [70] 【Y820】B(右側) 位置1ストッパー 行 異常表示; [71] 【Y821】B(右側) 位置2ストッパー戻 異常表示; [72] 【Y821】B(右側) 位置2ストッパー行 異常表示; [73] 【Y822】B(右側) 位置3ストッパー戻 異常表示; [74] 【Y822】B(右側) 位置3ストッパー行 異常表示; [75] 【Y823】B(右側) 位置4ストッパー戻 異常表示; [76] 【Y823】B(右側) 位置4ストッパー行 異常表示; [77] 【Y824】B(右側) 位置5ストッパー戻 異常表示; [78] 【Y824】B(右側) 位置5ストッパー行 異常表示; [79] 【Y825】B(右側) 位置6ストッパー戻 異常表示; [80] 【Y825】B(右側) 位置6ストッパー行 異常表示; [81] 【Y826】B(右側) ストックフォルダターン戻 異常表示; [82] 【Y827】B(右側) ストックフォルダターン行 異常表示; [83] 【Y828】B(右側) NG1仕分け 戻 異常表示; [84] 【Y829】B(右側) NG1仕分け 行 異常表示; [85] 【Y1200】空コンテナ送り 戻 異常表示; [86] 【Y1201】空コンテナ送り 行 異常表示; [87] 【Y1202】段バラシ爪 戻 異常表示; [88] 【Y1203】段バラシ爪 行 異常表示; [89] 【Y1204】コンテナ排出 戻 異常表示; [90] 【Y1205】コンテナ排出 行 異常表示; [91] Output_Share_Error_M[7] 異常表示; [92] 【Y1207】箱入れチャック 行 異常表示; [93] 【Y1208】コンテナ仕分けストッパー 戻 異常表示; [94] 【Y1209】コンテナ仕分けストッパー 行 異常表示; [95] 【Y1210】コンテナ仕分け送り 戻 異常表示; [96] Output_Share_Error_M[12] 異常表示; [97] 【Y1300】A(左側) コンベア受渡送り戻 異常表示; [98] 【Y1301】A(左側) コンベア受渡送り行 異常表示; [99] 【Y1302】B(右側) コンベア受渡送り戻 異常表示; [100] 【Y1303】B(右側) コンベア受渡送り行 異常表示; [101] ST1 搬送ワーク不一致; [102] ST2 搬送ワーク不一致; [103] ST3 搬送ワーク不一致; [104] ST4 搬送ワーク不一致; [105] ST5 搬送ワーク不一致; [106] ST6 搬送ワーク不一致; [107] ST7 搬送ワーク不一致; [108] A(左側) ST1 FH測定時間超過; [109] A(左側) ST1 FH異常; [110] A(左側) ST5 FH異常; [111] B(右側) ST1 FH異常; [112] B(右側) ST5 FH異常; [113] A(左側) ST1 FH判定OK; [114] A(左側) ST1 FH判定NG1; [115] A(左側) ST1 FH判定NG2; [116] A(左側) ST1 検査前ワーク不一致; [117] A(左側) ST5 FH測定時間超過; [118] A(左側) ST5 FH判定OK; [119] A(左側) ST5 FH判定NG1; [120] A(左側) ST5 FH判定NG2; [121] A(左側) ST5 検査前ワーク不一致 *)
    HMI_Error_WorkSample : ARRAY[0..1] OF BOOL;  (* #HMI 再開前のワーク不一致; [0] A(左側) ST1; [1] A(左側) ST5 *)
    Error_ST1_A_Timeout : BOOL;  (* FHタイムアウト（非保持） *)
    Error_ST5_A_Timeout : BOOL;  (* FHタイムアウト（非保持） *)
    TimerQ_In_Sen_Work_A_Pos_07 : BOOL;  (* 【X209】A(左側)ワーク位置7 *)
    TimerQ_In_Sen_NG2_Tray_B_Full : BOOL;  (* 【X412】B(右側) NG2トレイ満杯停止 *)
    Retry : ARRAY[0..99] OF BOOL;
    Stm_A_Rev1_Axis000_Power_Error : BOOL;
    Stm_A_Rev_Axis000_MoveError : BOOL;
    RCON1_3_Error : BOOL;
    RCON1_3_Error_Clear : BOOL;
    RCON1_3_IN_Alarm : BOOL;
    RCON1_3_IN_EmergencyStop : BOOL;
    TimerQ_In_Sen_NG2_Tray_A_Full : BOOL;
    RCON1_5_Error : BOOL;
    RCON1_5_Error_Clear : BOOL;
    Auto_Com_Start : BOOL;  (* 共通ユニット自動運転開始 *)
    Destacker_Error : BOOL;  (* 方向・1段目確認異常 *)
    Error_Destacker_M : ARRAY[0..99] OF Bool;  (* 段バラシエラー： *)
END_VAR
VAR
    _p1 : BOOL;
    _p2 : BOOL;
    _p3 : BOOL;
    _p4 : BOOL;
    _p5 : BOOL;
    _p6 : BOOL;
    _p7 : BOOL;
    _p8 : BOOL;
    _p9 : BOOL;
    _p10 : BOOL;
    _p11 : BOOL;
    _p12 : BOOL;
    _p13 : BOOL;
    _p14 : BOOL;
    _p15 : BOOL;
    _p16 : BOOL;
    _p17 : BOOL;
    _p18 : BOOL;
    _p19 : BOOL;
    _p20 : BOOL;
    _p21 : BOOL;
    _p22 : BOOL;
    _p23 : BOOL;
    _p24 : BOOL;
    _e25 : R_TRIG;
    _e26 : R_TRIG;
    _e27 : R_TRIG;
    _e28 : R_TRIG;
    _e29 : R_TRIG;
    _e30 : R_TRIG;
    _e31 : R_TRIG;
    _e32 : R_TRIG;
    _e33 : R_TRIG;
    _e34 : R_TRIG;
    _p35 : BOOL;
    _p36 : BOOL;
    _p37 : BOOL;
    _e38 : R_TRIG;
    _e39 : R_TRIG;
    _e40 : R_TRIG;
    _e41 : R_TRIG;
    _e42 : R_TRIG;
    _e43 : R_TRIG;
    _e44 : R_TRIG;
    _e45 : R_TRIG;
    _e46 : R_TRIG;
    _e47 : R_TRIG;
    _p48 : BOOL;
END_VAR

(* Section Initial_初期化処理: ladder, written here as Structured Text *)

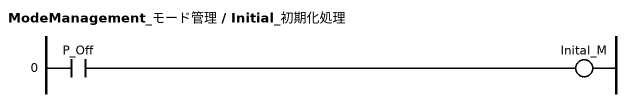
(* Rung 0 *)
Inital_M := P_Off;

(* Section Origin_原点復帰: ladder, written here as Structured Text *)

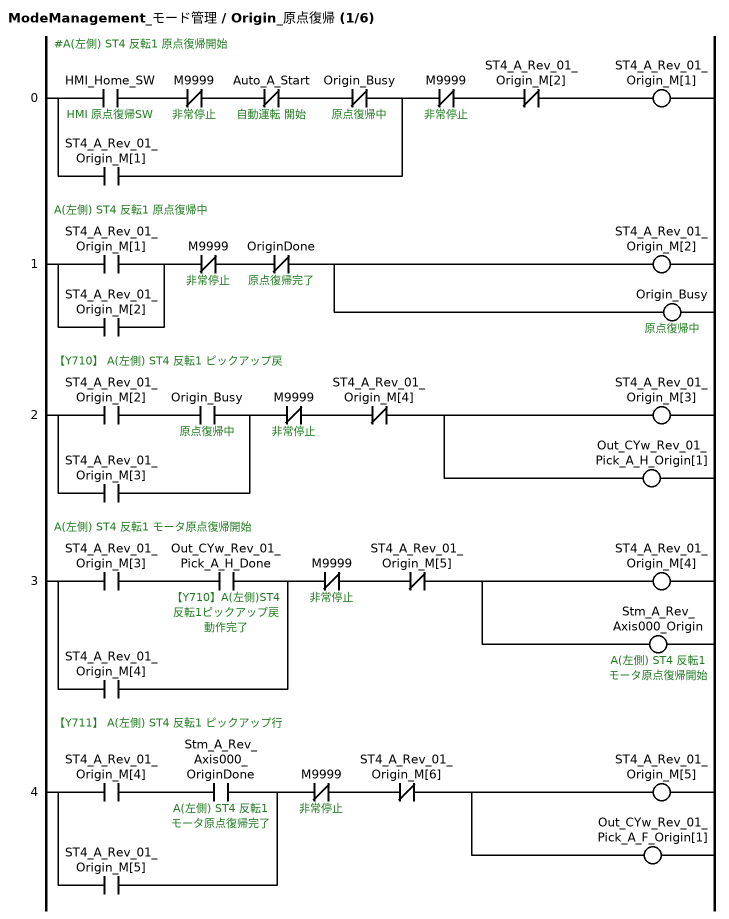
(* Rung 0: #A(左側) ST4 反転1 原点復帰開始 *)
ST4_A_Rev_01_Origin_M[1] := ((HMI_Home_SW AND NOT M9999 AND NOT Auto_A_Start AND NOT Origin_Busy) OR ST4_A_Rev_01_Origin_M[1]) AND NOT M9999 AND NOT ST4_A_Rev_01_Origin_M[2];
(* Rung 1: A(左側) ST4 反転1 原点復帰中 *)
_p1 := (ST4_A_Rev_01_Origin_M[1] OR ST4_A_Rev_01_Origin_M[2]) AND NOT M9999 AND NOT OriginDone;
ST4_A_Rev_01_Origin_M[2] := _p1;
Origin_Busy := _p1;
(* Rung 2: 【Y710】 A(左側) ST4 反転1 ピックアップ戻 *)
_p2 := ((ST4_A_Rev_01_Origin_M[2] AND Origin_Busy) OR ST4_A_Rev_01_Origin_M[3]) AND NOT M9999 AND NOT ST4_A_Rev_01_Origin_M[4];
ST4_A_Rev_01_Origin_M[3] := _p2;
Out_CYw_Rev_01_Pick_A_H_Origin[1] := _p2;
(* Rung 3: A(左側) ST4 反転1 モータ原点復帰開始 *)
_p3 := ((ST4_A_Rev_01_Origin_M[3] AND Out_CYw_Rev_01_Pick_A_H_Done) OR ST4_A_Rev_01_Origin_M[4]) AND NOT M9999 AND NOT ST4_A_Rev_01_Origin_M[5];
ST4_A_Rev_01_Origin_M[4] := _p3;
Stm_A_Rev_Axis000_Origin := _p3;
(* Rung 4: 【Y711】 A(左側) ST4 反転1 ピックアップ行 *)
_p4 := ((ST4_A_Rev_01_Origin_M[4] AND Stm_A_Rev_Axis000_OriginDone) OR ST4_A_Rev_01_Origin_M[5]) AND NOT M9999 AND NOT ST4_A_Rev_01_Origin_M[6];
ST4_A_Rev_01_Origin_M[5] := _p4;
Out_CYw_Rev_01_Pick_A_F_Origin[1] := _p4;

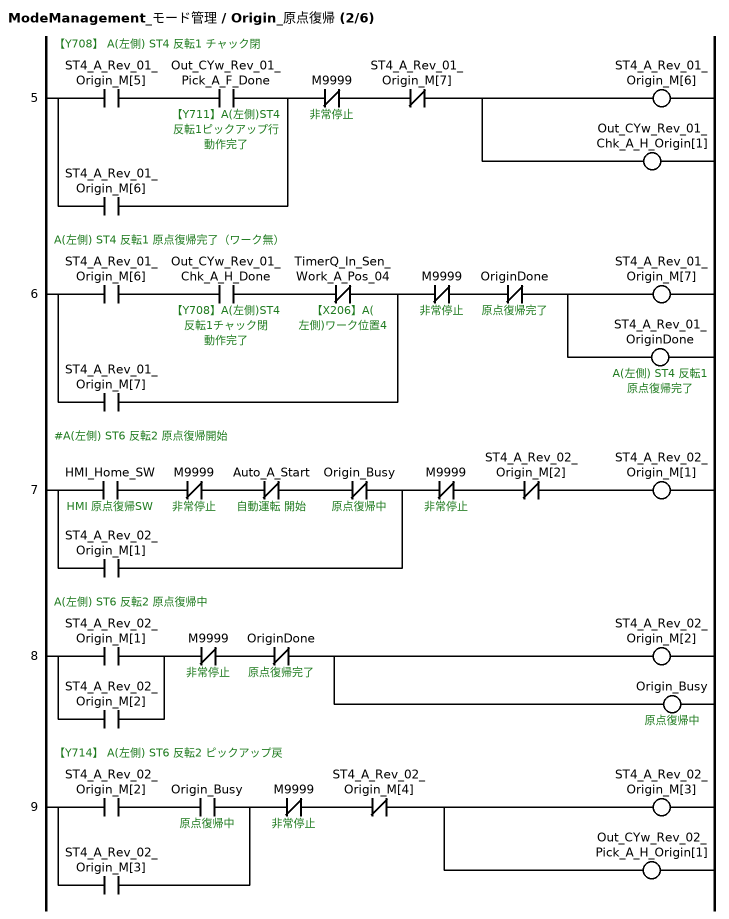
(* Rung 5: 【Y708】 A(左側) ST4 反転1 チャック閉 *)
_p5 := ((ST4_A_Rev_01_Origin_M[5] AND Out_CYw_Rev_01_Pick_A_F_Done) OR ST4_A_Rev_01_Origin_M[6]) AND NOT M9999 AND NOT ST4_A_Rev_01_Origin_M[7];
ST4_A_Rev_01_Origin_M[6] := _p5;
Out_CYw_Rev_01_Chk_A_H_Origin[1] := _p5;
(* Rung 6: A(左側) ST4 反転1 原点復帰完了（ワーク無） *)
_p6 := ((ST4_A_Rev_01_Origin_M[6] AND Out_CYw_Rev_01_Chk_A_H_Done AND NOT TimerQ_In_Sen_Work_A_Pos_04) OR ST4_A_Rev_01_Origin_M[7]) AND NOT M9999 AND NOT OriginDone;
ST4_A_Rev_01_Origin_M[7] := _p6;
ST4_A_Rev_01_OriginDone := _p6;
(* Rung 7: #A(左側) ST6 反転2 原点復帰開始 *)
ST4_A_Rev_02_Origin_M[1] := ((HMI_Home_SW AND NOT M9999 AND NOT Auto_A_Start AND NOT Origin_Busy) OR ST4_A_Rev_02_Origin_M[1]) AND NOT M9999 AND NOT ST4_A_Rev_02_Origin_M[2];
(* Rung 8: A(左側) ST6 反転2 原点復帰中 *)
_p7 := (ST4_A_Rev_02_Origin_M[1] OR ST4_A_Rev_02_Origin_M[2]) AND NOT M9999 AND NOT OriginDone;
ST4_A_Rev_02_Origin_M[2] := _p7;
Origin_Busy := _p7;
(* Rung 9: 【Y714】 A(左側) ST6 反転2 ピックアップ戻 *)
_p8 := ((ST4_A_Rev_02_Origin_M[2] AND Origin_Busy) OR ST4_A_Rev_02_Origin_M[3]) AND NOT M9999 AND NOT ST4_A_Rev_02_Origin_M[4];
ST4_A_Rev_02_Origin_M[3] := _p8;
Out_CYw_Rev_02_Pick_A_H_Origin[1] := _p8;

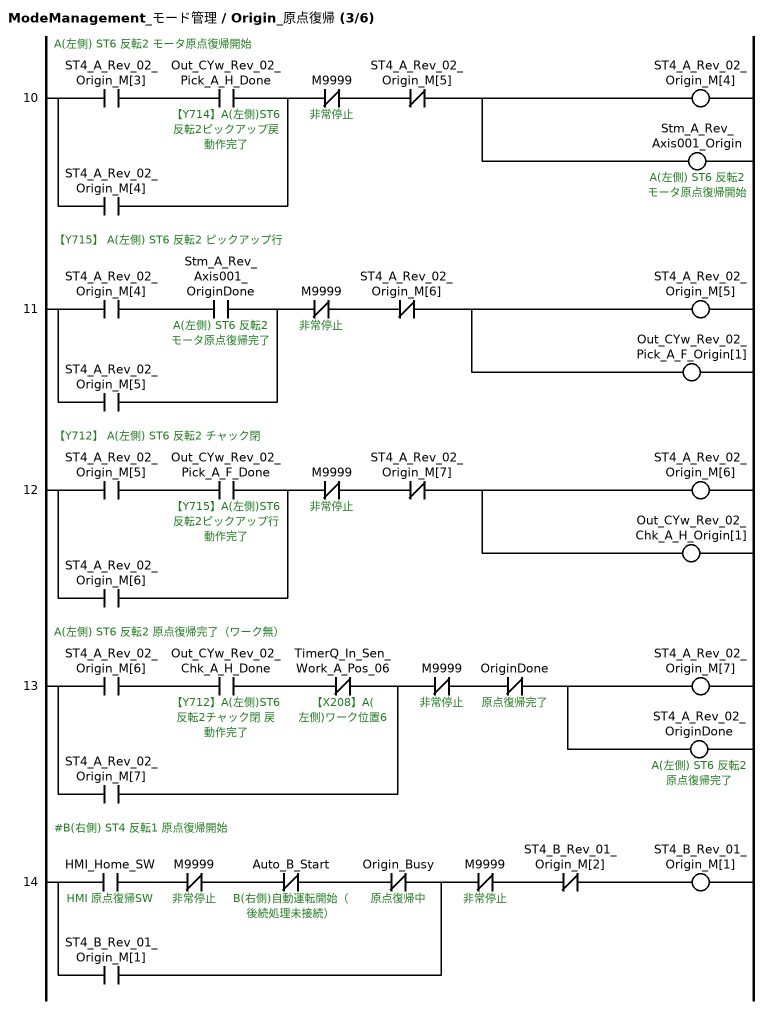
(* Rung 10: A(左側) ST6 反転2 モータ原点復帰開始 *)
_p9 := ((ST4_A_Rev_02_Origin_M[3] AND Out_CYw_Rev_02_Pick_A_H_Done) OR ST4_A_Rev_02_Origin_M[4]) AND NOT M9999 AND NOT ST4_A_Rev_02_Origin_M[5];
ST4_A_Rev_02_Origin_M[4] := _p9;
Stm_A_Rev_Axis001_Origin := _p9;
(* Rung 11: 【Y715】 A(左側) ST6 反転2 ピックアップ行 *)
_p10 := ((ST4_A_Rev_02_Origin_M[4] AND Stm_A_Rev_Axis001_OriginDone) OR ST4_A_Rev_02_Origin_M[5]) AND NOT M9999 AND NOT ST4_A_Rev_02_Origin_M[6];
ST4_A_Rev_02_Origin_M[5] := _p10;
Out_CYw_Rev_02_Pick_A_F_Origin[1] := _p10;
(* Rung 12: 【Y712】 A(左側) ST6 反転2 チャック閉 *)
_p11 := ((ST4_A_Rev_02_Origin_M[5] AND Out_CYw_Rev_02_Pick_A_F_Done) OR ST4_A_Rev_02_Origin_M[6]) AND NOT M9999 AND NOT ST4_A_Rev_02_Origin_M[7];
ST4_A_Rev_02_Origin_M[6] := _p11;
Out_CYw_Rev_02_Chk_A_H_Origin[1] := _p11;
(* Rung 13: A(左側) ST6 反転2 原点復帰完了（ワーク無） *)
_p12 := ((ST4_A_Rev_02_Origin_M[6] AND Out_CYw_Rev_02_Chk_A_H_Done AND NOT TimerQ_In_Sen_Work_A_Pos_06) OR ST4_A_Rev_02_Origin_M[7]) AND NOT M9999 AND NOT OriginDone;
ST4_A_Rev_02_Origin_M[7] := _p12;
ST4_A_Rev_02_OriginDone := _p12;
(* Rung 14: #B(右側) ST4 反転1 原点復帰開始 *)
ST4_B_Rev_01_Origin_M[1] := ((HMI_Home_SW AND NOT M9999 AND NOT Auto_B_Start AND NOT Origin_Busy) OR ST4_B_Rev_01_Origin_M[1]) AND NOT M9999 AND NOT ST4_B_Rev_01_Origin_M[2];

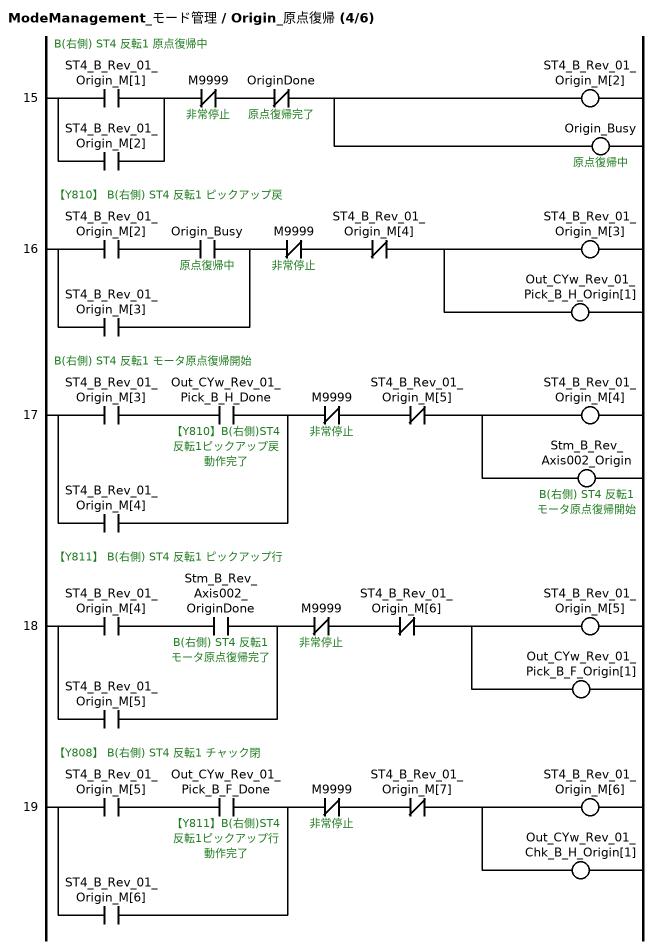
(* Rung 15: B(右側) ST4 反転1 原点復帰中 *)
_p13 := (ST4_B_Rev_01_Origin_M[1] OR ST4_B_Rev_01_Origin_M[2]) AND NOT M9999 AND NOT OriginDone;
ST4_B_Rev_01_Origin_M[2] := _p13;
Origin_Busy := _p13;
(* Rung 16: 【Y810】 B(右側) ST4 反転1 ピックアップ戻 *)
_p14 := ((ST4_B_Rev_01_Origin_M[2] AND Origin_Busy) OR ST4_B_Rev_01_Origin_M[3]) AND NOT M9999 AND NOT ST4_B_Rev_01_Origin_M[4];
ST4_B_Rev_01_Origin_M[3] := _p14;
Out_CYw_Rev_01_Pick_B_H_Origin[1] := _p14;
(* Rung 17: B(右側) ST4 反転1 モータ原点復帰開始 *)
_p15 := ((ST4_B_Rev_01_Origin_M[3] AND Out_CYw_Rev_01_Pick_B_H_Done) OR ST4_B_Rev_01_Origin_M[4]) AND NOT M9999 AND NOT ST4_B_Rev_01_Origin_M[5];
ST4_B_Rev_01_Origin_M[4] := _p15;
Stm_B_Rev_Axis002_Origin := _p15;
(* Rung 18: 【Y811】 B(右側) ST4 反転1 ピックアップ行 *)
_p16 := ((ST4_B_Rev_01_Origin_M[4] AND Stm_B_Rev_Axis002_OriginDone) OR ST4_B_Rev_01_Origin_M[5]) AND NOT M9999 AND NOT ST4_B_Rev_01_Origin_M[6];
ST4_B_Rev_01_Origin_M[5] := _p16;
Out_CYw_Rev_01_Pick_B_F_Origin[1] := _p16;
(* Rung 19: 【Y808】 B(右側) ST4 反転1 チャック閉 *)
_p17 := ((ST4_B_Rev_01_Origin_M[5] AND Out_CYw_Rev_01_Pick_B_F_Done) OR ST4_B_Rev_01_Origin_M[6]) AND NOT M9999 AND NOT ST4_B_Rev_01_Origin_M[7];
ST4_B_Rev_01_Origin_M[6] := _p17;
Out_CYw_Rev_01_Chk_B_H_Origin[1] := _p17;

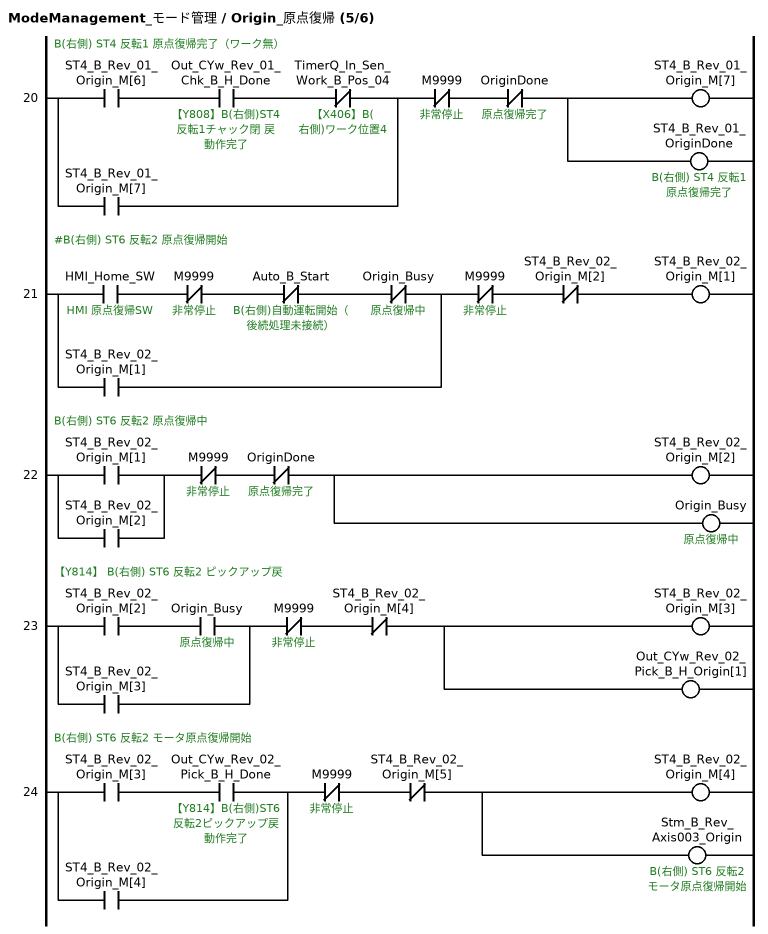
(* Rung 20: B(右側) ST4 反転1 原点復帰完了（ワーク無） *)
_p18 := ((ST4_B_Rev_01_Origin_M[6] AND Out_CYw_Rev_01_Chk_B_H_Done AND NOT TimerQ_In_Sen_Work_B_Pos_04) OR ST4_B_Rev_01_Origin_M[7]) AND NOT M9999 AND NOT OriginDone;
ST4_B_Rev_01_Origin_M[7] := _p18;
ST4_B_Rev_01_OriginDone := _p18;
(* Rung 21: #B(右側) ST6 反転2 原点復帰開始 *)
ST4_B_Rev_02_Origin_M[1] := ((HMI_Home_SW AND NOT M9999 AND NOT Auto_B_Start AND NOT Origin_Busy) OR ST4_B_Rev_02_Origin_M[1]) AND NOT M9999 AND NOT ST4_B_Rev_02_Origin_M[2];
(* Rung 22: B(右側) ST6 反転2 原点復帰中 *)
_p19 := (ST4_B_Rev_02_Origin_M[1] OR ST4_B_Rev_02_Origin_M[2]) AND NOT M9999 AND NOT OriginDone;
ST4_B_Rev_02_Origin_M[2] := _p19;
Origin_Busy := _p19;
(* Rung 23: 【Y814】 B(右側) ST6 反転2 ピックアップ戻 *)
_p20 := ((ST4_B_Rev_02_Origin_M[2] AND Origin_Busy) OR ST4_B_Rev_02_Origin_M[3]) AND NOT M9999 AND NOT ST4_B_Rev_02_Origin_M[4];
ST4_B_Rev_02_Origin_M[3] := _p20;
Out_CYw_Rev_02_Pick_B_H_Origin[1] := _p20;
(* Rung 24: B(右側) ST6 反転2 モータ原点復帰開始 *)
_p21 := ((ST4_B_Rev_02_Origin_M[3] AND Out_CYw_Rev_02_Pick_B_H_Done) OR ST4_B_Rev_02_Origin_M[4]) AND NOT M9999 AND NOT ST4_B_Rev_02_Origin_M[5];
ST4_B_Rev_02_Origin_M[4] := _p21;
Stm_B_Rev_Axis003_Origin := _p21;

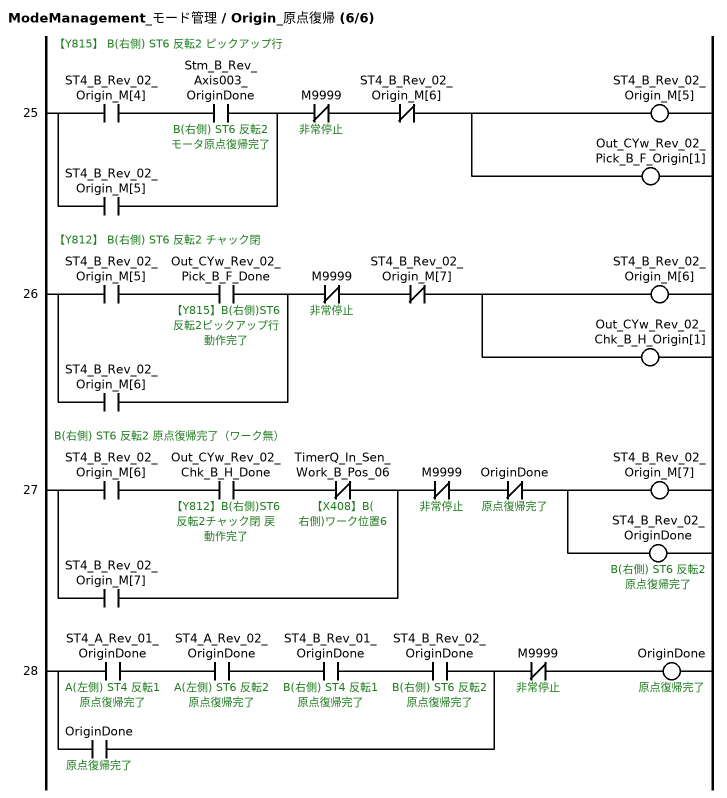
(* Rung 25: 【Y815】 B(右側) ST6 反転2 ピックアップ行 *)
_p22 := ((ST4_B_Rev_02_Origin_M[4] AND Stm_B_Rev_Axis003_OriginDone) OR ST4_B_Rev_02_Origin_M[5]) AND NOT M9999 AND NOT ST4_B_Rev_02_Origin_M[6];
ST4_B_Rev_02_Origin_M[5] := _p22;
Out_CYw_Rev_02_Pick_B_F_Origin[1] := _p22;
(* Rung 26: 【Y812】 B(右側) ST6 反転2 チャック閉 *)
_p23 := ((ST4_B_Rev_02_Origin_M[5] AND Out_CYw_Rev_02_Pick_B_F_Done) OR ST4_B_Rev_02_Origin_M[6]) AND NOT M9999 AND NOT ST4_B_Rev_02_Origin_M[7];
ST4_B_Rev_02_Origin_M[6] := _p23;
Out_CYw_Rev_02_Chk_B_H_Origin[1] := _p23;
(* Rung 27: B(右側) ST6 反転2 原点復帰完了（ワーク無） *)
_p24 := ((ST4_B_Rev_02_Origin_M[6] AND Out_CYw_Rev_02_Chk_B_H_Done AND NOT TimerQ_In_Sen_Work_B_Pos_06) OR ST4_B_Rev_02_Origin_M[7]) AND NOT M9999 AND NOT OriginDone;
ST4_B_Rev_02_Origin_M[7] := _p24;
ST4_B_Rev_02_OriginDone := _p24;
(* Rung 28 *)
OriginDone := ((ST4_A_Rev_01_OriginDone AND ST4_A_Rev_02_OriginDone AND ST4_B_Rev_01_OriginDone AND ST4_B_Rev_02_OriginDone) OR OriginDone) AND NOT M9999;

(* Section DummyCheck_ダミーチェック: ladder, written here as Structured Text *)

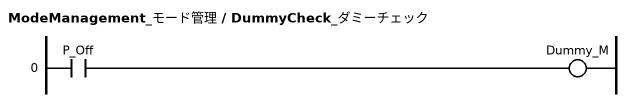
(* Rung 0 *)
Dummy_M := P_Off;

(* Section AutoMode_自動運転: ladder, written here as Structured Text *)

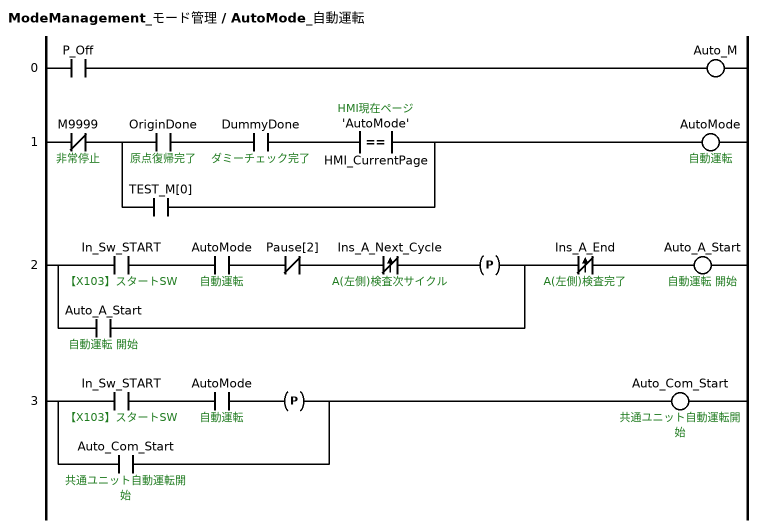
(* Rung 0 *)
Auto_M := P_Off;
(* Rung 1 *)
AutoMode := NOT M9999 AND ((OriginDone AND DummyDone AND ('AutoMode' = HMI_CurrentPage)) OR TEST_M[0]);
(* Rung 2 *)
_e25(CLK := Ins_A_Next_Cycle);
_e26(CLK := In_Sw_START AND AutoMode AND NOT Pause[2] AND NOT _e25.Q);
_e27(CLK := Ins_A_End);
Auto_A_Start := (_e26.Q OR Auto_A_Start) AND NOT _e27.Q;
(* Rung 3 *)
_e28(CLK := In_Sw_START AND AutoMode);
Auto_Com_Start := _e28.Q OR Auto_Com_Start;

(* Section Manual_手動運転: ladder, written here as Structured Text *)

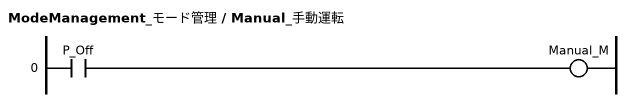
(* Rung 0 *)
Manual_M := P_Off;

(* Section Setting_設定: ladder, written here as Structured Text *)

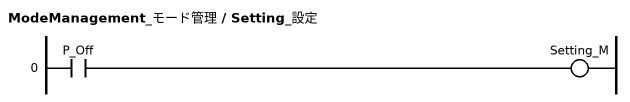
(* Rung 0 *)
Setting_M := P_Off;

(* Section Error_エラー処理: ladder, written here as Structured Text *)

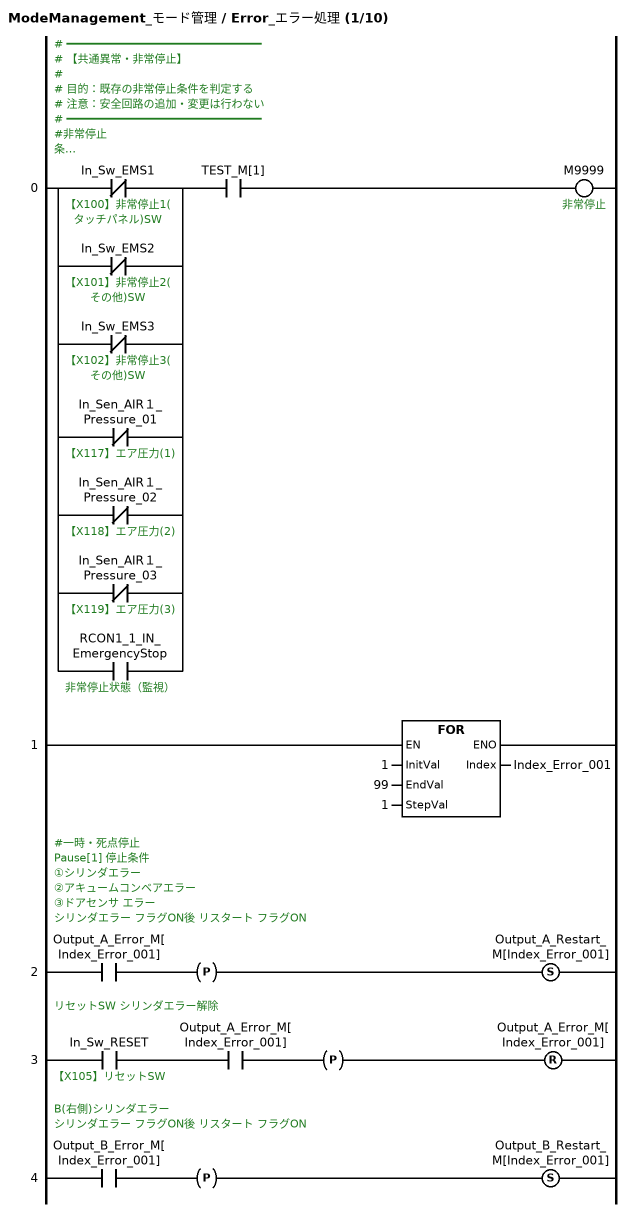
(* Rung 0: # ━━━━━━━━━━━━━━━━━━━━━━━━━━━━━━ / # 【共通異常・非常停止】 / # / # 目的：既存の非常停止条件を判定する / # 注意：安全回路の追加・変更は行わない / # ━━━━━━━━━━━━━━━━━━━━━━━━━━━━━━ / #非常停止 / 条件 / ①非常停止SW ON / ②エア圧力 低下 *)
M9999 := (NOT In_Sw_EMS1 OR NOT In_Sw_EMS2 OR NOT In_Sw_EMS3 OR NOT In_Sen_AIR１_Pressure_01 OR NOT In_Sen_AIR１_Pressure_02 OR NOT In_Sen_AIR１_Pressure_03 OR RCON1_1_IN_EmergencyStop) AND TEST_M[1];
(* Rung 1 *)
Index_Error_001 := FOR(InitVal := 1, EndVal := 99, StepVal := 1);
(* Rung 2: #一時・死点停止 / Pause[1] 停止条件 / ①シリンダエラー / ②アキュームコンベアエラー / ③ドアセンサ エラー / シリンダエラー フラグON後 リスタート フラグON *)
_e29(CLK := Output_A_Error_M[Index_Error_001]);
IF _e29.Q THEN Output_A_Restart_M[Index_Error_001] := TRUE; END_IF;
(* Rung 3: リセットSW シリンダエラー解除 *)
_e30(CLK := In_Sw_RESET AND Output_A_Error_M[Index_Error_001]);
IF _e30.Q THEN Output_A_Error_M[Index_Error_001] := FALSE; END_IF;
(* Rung 4: B(右側)シリンダエラー / シリンダエラー フラグON後 リスタート フラグON *)
_e31(CLK := Output_B_Error_M[Index_Error_001]);
IF _e31.Q THEN Output_B_Restart_M[Index_Error_001] := TRUE; END_IF;

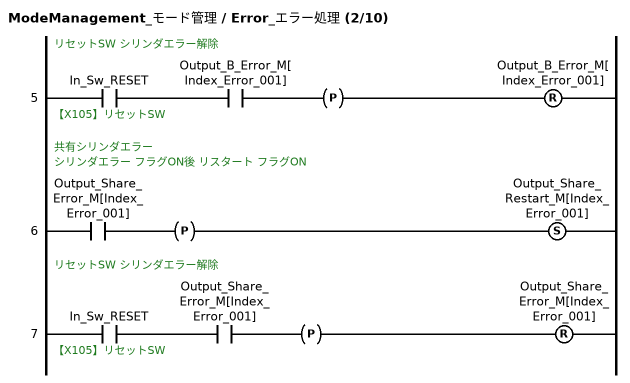
(* Rung 5: リセットSW シリンダエラー解除 *)
_e32(CLK := In_Sw_RESET AND Output_B_Error_M[Index_Error_001]);
IF _e32.Q THEN Output_B_Error_M[Index_Error_001] := FALSE; END_IF;
(* Rung 6: 共有シリンダエラー / シリンダエラー フラグON後 リスタート フラグON *)
_e33(CLK := Output_Share_Error_M[Index_Error_001]);
IF _e33.Q THEN Output_Share_Restart_M[Index_Error_001] := TRUE; END_IF;
(* Rung 7: リセットSW シリンダエラー解除 *)
_e34(CLK := In_Sw_RESET AND Output_Share_Error_M[Index_Error_001]);
IF _e34.Q THEN Output_Share_Error_M[Index_Error_001] := FALSE; END_IF;

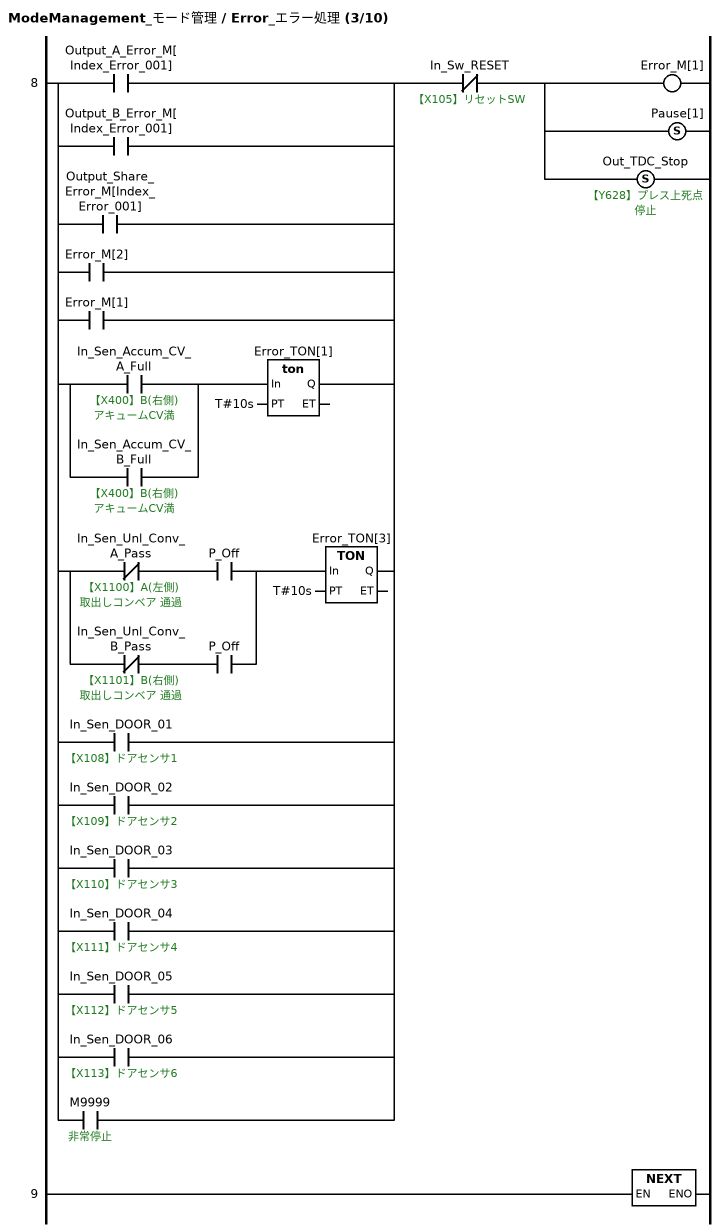
(* Rung 8 *)
Error_TON[1](In := In_Sen_Accum_CV_A_Full OR In_Sen_Accum_CV_B_Full, PT := T#10s);
_p35 := Error_TON[1].Q;
Error_TON[3](In := (NOT In_Sen_Unl_Conv_A_Pass AND P_Off) OR (NOT In_Sen_Unl_Conv_B_Pass AND P_Off), PT := T#10s);
_p36 := (Output_A_Error_M[Index_Error_001] OR Output_B_Error_M[Index_Error_001] OR Output_Share_Error_M[Index_Error_001] OR Error_M[2] OR Error_M[1] OR _p35 OR Error_TON[3].Q OR In_Sen_DOOR_01 OR In_Sen_DOOR_02 OR In_Sen_DOOR_03 OR In_Sen_DOOR_04 OR In_Sen_DOOR_05 OR In_Sen_DOOR_06 OR M9999) AND NOT In_Sw_RESET;
Error_M[1] := _p36;
IF _p36 THEN
    Pause[1] := TRUE;
    Out_TDC_Stop := TRUE;
END_IF;
(* Rung 9 *)
NEXT();

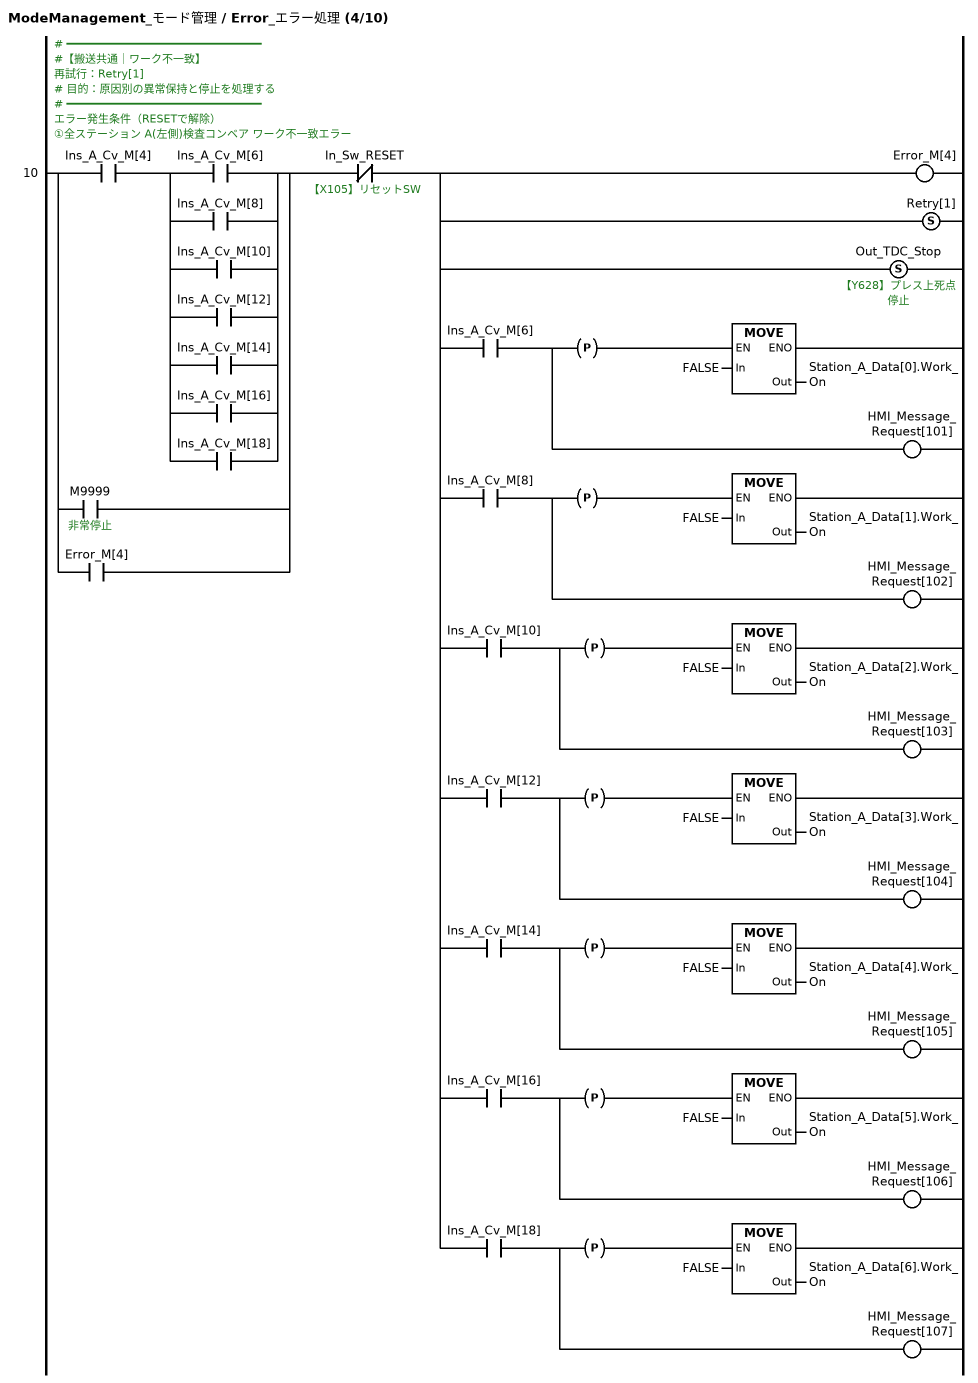
(* Rung 10: # ━━━━━━━━━━━━━━━━━━━━━━━━━━━━━━ / #【搬送共通｜ワーク不一致】 / 再試行：Retry[1] / # 目的：原因別の異常保持と停止を処理する / # ━━━━━━━━━━━━━━━━━━━━━━━━━━━━━━ / エラー発生条件（RESETで解除） / ①全ステーション A(左側)検査コンベア ワーク不一致エラー *)
_p37 := ((Ins_A_Cv_M[4] AND (Ins_A_Cv_M[6] OR Ins_A_Cv_M[8] OR Ins_A_Cv_M[10] OR Ins_A_Cv_M[12] OR Ins_A_Cv_M[14] OR Ins_A_Cv_M[16] OR Ins_A_Cv_M[18])) OR M9999 OR Error_M[4]) AND NOT In_Sw_RESET;
Error_M[4] := _p37;
IF _p37 THEN
    Retry[1] := TRUE;
    Out_TDC_Stop := TRUE;
END_IF;
_e38(CLK := _p37 AND Ins_A_Cv_M[6]);
IF _e38.Q THEN Station_A_Data[0].Work_On := FALSE; END_IF;
HMI_Message_Request[101] := _p37 AND Ins_A_Cv_M[6];
_e39(CLK := _p37 AND Ins_A_Cv_M[8]);
IF _e39.Q THEN Station_A_Data[1].Work_On := FALSE; END_IF;
HMI_Message_Request[102] := _p37 AND Ins_A_Cv_M[8];
_e40(CLK := _p37 AND Ins_A_Cv_M[10]);
IF _e40.Q THEN Station_A_Data[2].Work_On := FALSE; END_IF;
HMI_Message_Request[103] := _p37 AND Ins_A_Cv_M[10];
_e41(CLK := _p37 AND Ins_A_Cv_M[12]);
IF _e41.Q THEN Station_A_Data[3].Work_On := FALSE; END_IF;
HMI_Message_Request[104] := _p37 AND Ins_A_Cv_M[12];
_e42(CLK := _p37 AND Ins_A_Cv_M[14]);
IF _e42.Q THEN Station_A_Data[4].Work_On := FALSE; END_IF;
HMI_Message_Request[105] := _p37 AND Ins_A_Cv_M[14];
_e43(CLK := _p37 AND Ins_A_Cv_M[16]);
IF _e43.Q THEN Station_A_Data[5].Work_On := FALSE; END_IF;
HMI_Message_Request[106] := _p37 AND Ins_A_Cv_M[16];
_e44(CLK := _p37 AND Ins_A_Cv_M[18]);
IF _e44.Q THEN Station_A_Data[6].Work_On := FALSE; END_IF;
HMI_Message_Request[107] := _p37 AND Ins_A_Cv_M[18];

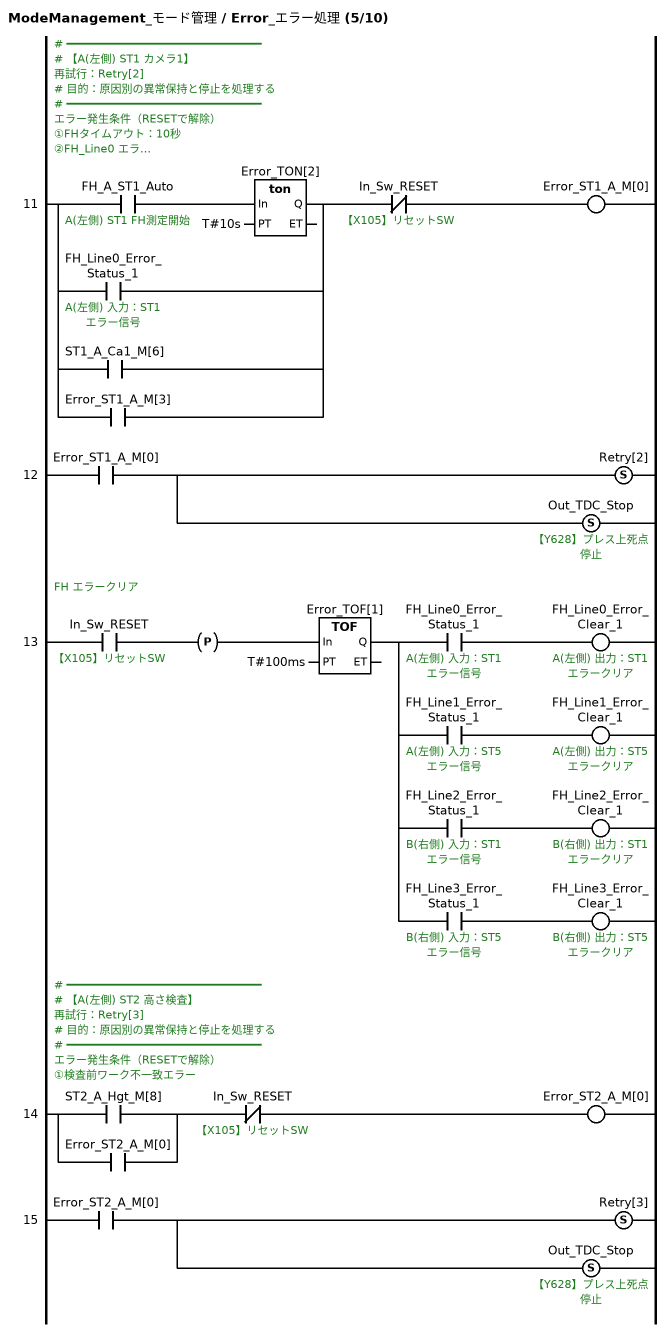
(* Rung 11: # ━━━━━━━━━━━━━━━━━━━━━━━━━━━━━━ / # 【A(左側) ST1 カメラ1】 / 再試行：Retry[2] / # 目的：原因別の異常保持と停止を処理する / # ━━━━━━━━━━━━━━━━━━━━━━━━━━━━━━ / エラー発生条件（RESETで解除） / ①FHタイムアウト：10秒 / ②FH_Line0 エラー / ③検査前ワーク不一致 *)
Error_TON[2](In := FH_A_ST1_Auto, PT := T#10s);
Error_ST1_A_M[0] := (Error_TON[2].Q OR FH_Line0_Error_Status_1 OR ST1_A_Ca1_M[6] OR Error_ST1_A_M[3]) AND NOT In_Sw_RESET;
(* Rung 12 *)
IF Error_ST1_A_M[0] THEN
    Retry[2] := TRUE;
    Out_TDC_Stop := TRUE;
END_IF;
(* Rung 13: FH エラークリア *)
_e45(CLK := In_Sw_RESET);
Error_TOF[1](In := _e45.Q, PT := T#100ms);
FH_Line0_Error_Clear_1 := Error_TOF[1].Q AND FH_Line0_Error_Status_1;
FH_Line1_Error_Clear_1 := Error_TOF[1].Q AND FH_Line1_Error_Status_1;
FH_Line2_Error_Clear_1 := Error_TOF[1].Q AND FH_Line2_Error_Status_1;
FH_Line3_Error_Clear_1 := Error_TOF[1].Q AND FH_Line3_Error_Status_1;
(* Rung 14: # ━━━━━━━━━━━━━━━━━━━━━━━━━━━━━━ / # 【A(左側) ST2 高さ検査】 / 再試行：Retry[3] / # 目的：原因別の異常保持と停止を処理する / # ━━━━━━━━━━━━━━━━━━━━━━━━━━━━━━ / エラー発生条件（RESETで解除） / ①検査前ワーク不一致エラー *)
Error_ST2_A_M[0] := (ST2_A_Hgt_M[8] OR Error_ST2_A_M[0]) AND NOT In_Sw_RESET;
(* Rung 15 *)
IF Error_ST2_A_M[0] THEN
    Retry[3] := TRUE;
    Out_TDC_Stop := TRUE;
END_IF;

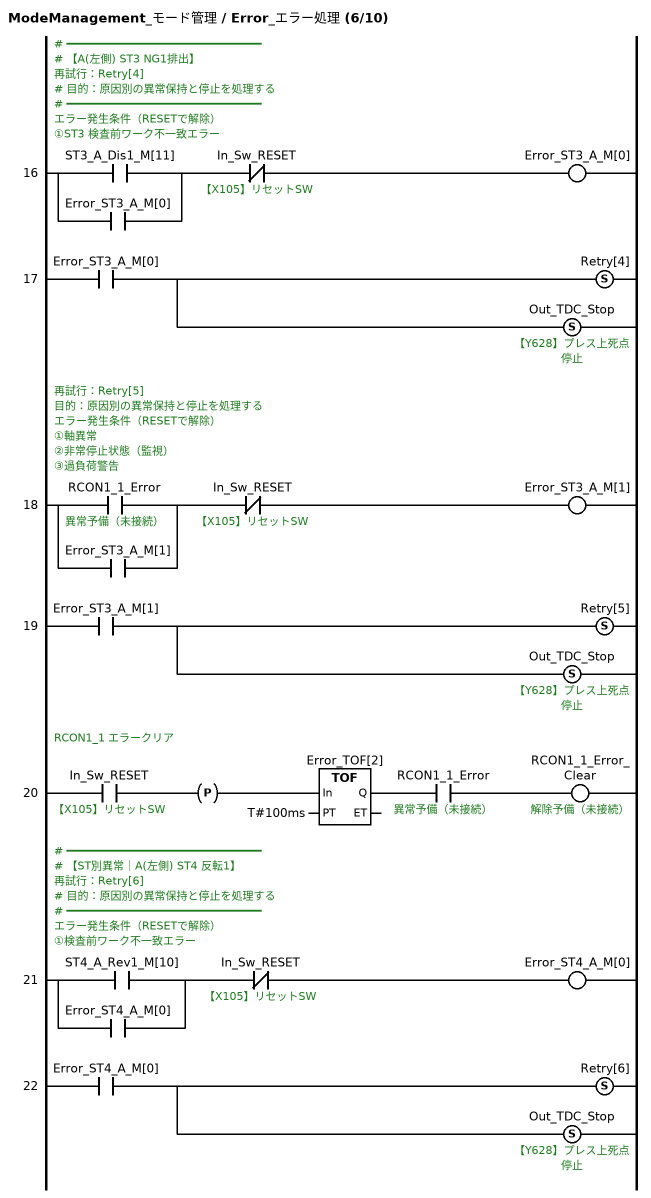
(* Rung 16: # ━━━━━━━━━━━━━━━━━━━━━━━━━━━━━━ / # 【A(左側) ST3 NG1排出】 / 再試行：Retry[4] / # 目的：原因別の異常保持と停止を処理する / # ━━━━━━━━━━━━━━━━━━━━━━━━━━━━━━ / エラー発生条件（RESETで解除） / ①ST3 検査前ワーク不一致エラー *)
Error_ST3_A_M[0] := (ST3_A_Dis1_M[11] OR Error_ST3_A_M[0]) AND NOT In_Sw_RESET;
(* Rung 17 *)
IF Error_ST3_A_M[0] THEN
    Retry[4] := TRUE;
    Out_TDC_Stop := TRUE;
END_IF;
(* Rung 18: 再試行：Retry[5] / 目的：原因別の異常保持と停止を処理する / エラー発生条件（RESETで解除） / ①軸異常 / ②非常停止状態（監視） / ③過負荷警告 *)
Error_ST3_A_M[1] := (RCON1_1_Error OR Error_ST3_A_M[1]) AND NOT In_Sw_RESET;
(* Rung 19 *)
IF Error_ST3_A_M[1] THEN
    Retry[5] := TRUE;
    Out_TDC_Stop := TRUE;
END_IF;
(* Rung 20: RCON1_1 エラークリア *)
_e46(CLK := In_Sw_RESET);
Error_TOF[2](In := _e46.Q, PT := T#100ms);
RCON1_1_Error_Clear := Error_TOF[2].Q AND RCON1_1_Error;
(* Rung 21: # ━━━━━━━━━━━━━━━━━━━━━━━━━━━━━━ / # 【ST別異常｜A(左側) ST4 反転1】 / 再試行：Retry[6] / # 目的：原因別の異常保持と停止を処理する / # ━━━━━━━━━━━━━━━━━━━━━━━━━━━━━━ / エラー発生条件（RESETで解除） / ①検査前ワーク不一致エラー *)
Error_ST4_A_M[0] := (ST4_A_Rev1_M[10] OR Error_ST4_A_M[0]) AND NOT In_Sw_RESET;
(* Rung 22 *)
IF Error_ST4_A_M[0] THEN
    Retry[6] := TRUE;
    Out_TDC_Stop := TRUE;
END_IF;

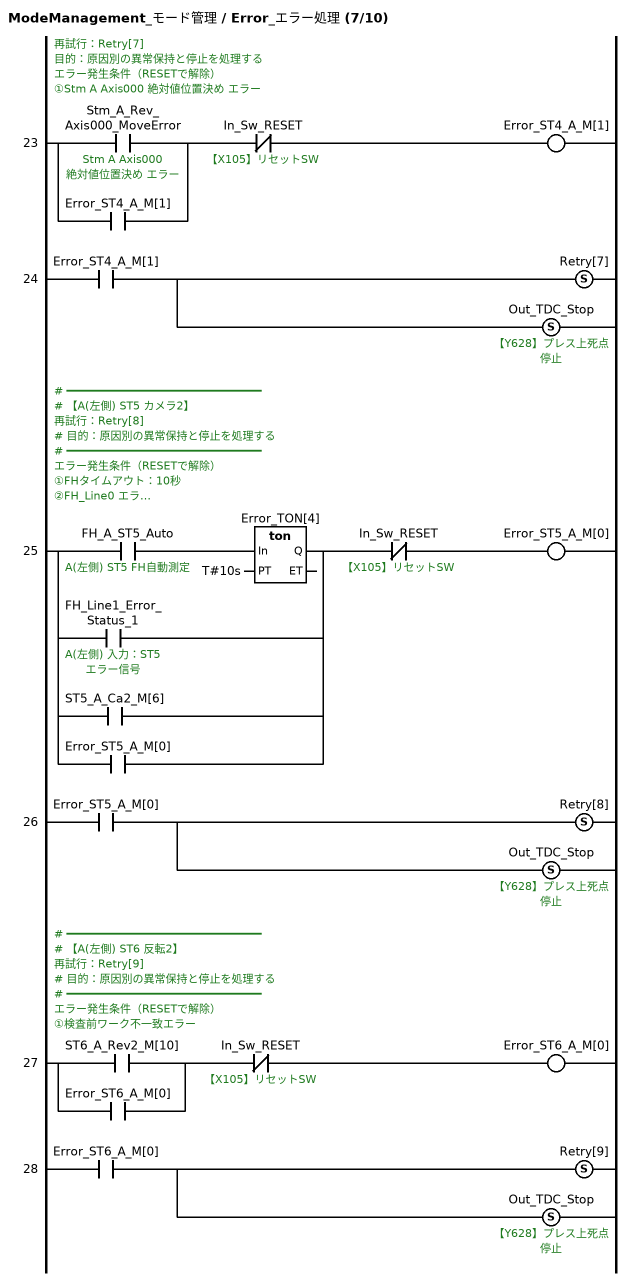
(* Rung 23: 再試行：Retry[7] / 目的：原因別の異常保持と停止を処理する / エラー発生条件（RESETで解除） / ①Stm A Axis000 絶対値位置決め エラー *)
Error_ST4_A_M[1] := (Stm_A_Rev_Axis000_MoveError OR Error_ST4_A_M[1]) AND NOT In_Sw_RESET;
(* Rung 24 *)
IF Error_ST4_A_M[1] THEN
    Retry[7] := TRUE;
    Out_TDC_Stop := TRUE;
END_IF;
(* Rung 25: # ━━━━━━━━━━━━━━━━━━━━━━━━━━━━━━ / # 【A(左側) ST5 カメラ2】 / 再試行：Retry[8] / # 目的：原因別の異常保持と停止を処理する / # ━━━━━━━━━━━━━━━━━━━━━━━━━━━━━━ / エラー発生条件（RESETで解除） / ①FHタイムアウト：10秒 / ②FH_Line0 エラー / ③検査前ワーク不一致 *)
Error_TON[4](In := FH_A_ST5_Auto, PT := T#10s);
Error_ST5_A_M[0] := (Error_TON[4].Q OR FH_Line1_Error_Status_1 OR ST5_A_Ca2_M[6] OR Error_ST5_A_M[0]) AND NOT In_Sw_RESET;
(* Rung 26 *)
IF Error_ST5_A_M[0] THEN
    Retry[8] := TRUE;
    Out_TDC_Stop := TRUE;
END_IF;
(* Rung 27: # ━━━━━━━━━━━━━━━━━━━━━━━━━━━━━━ / # 【A(左側) ST6 反転2】 / 再試行：Retry[9] / # 目的：原因別の異常保持と停止を処理する / # ━━━━━━━━━━━━━━━━━━━━━━━━━━━━━━ / エラー発生条件（RESETで解除） / ①検査前ワーク不一致エラー *)
Error_ST6_A_M[0] := (ST6_A_Rev2_M[10] OR Error_ST6_A_M[0]) AND NOT In_Sw_RESET;
(* Rung 28 *)
IF Error_ST6_A_M[0] THEN
    Retry[9] := TRUE;
    Out_TDC_Stop := TRUE;
END_IF;

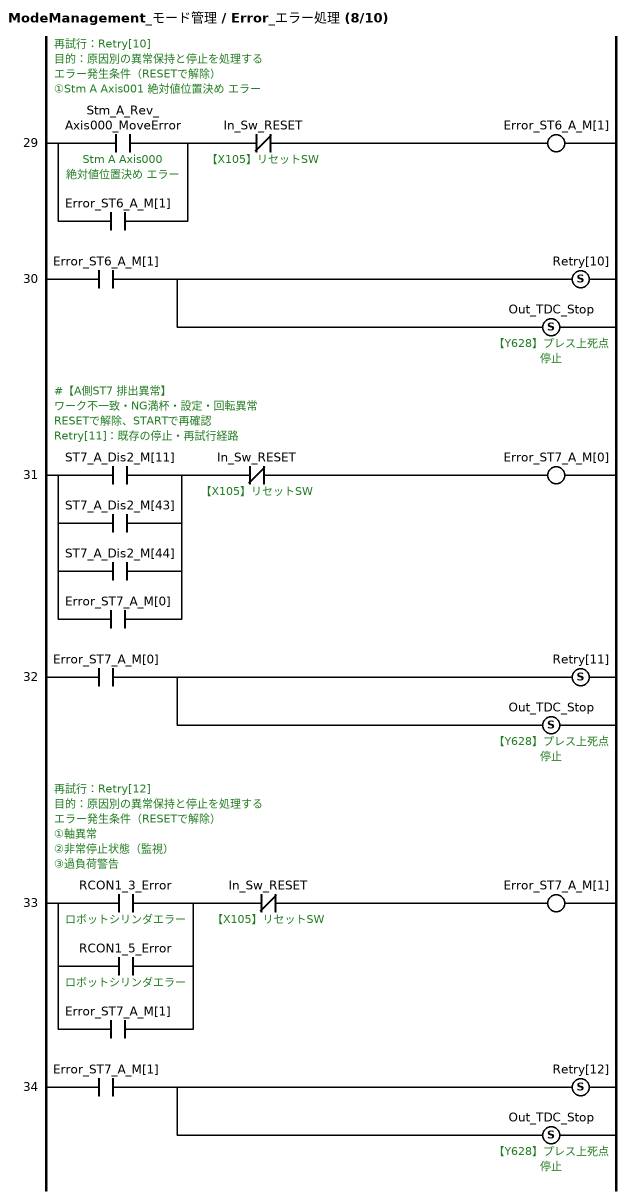
(* Rung 29: 再試行：Retry[10] / 目的：原因別の異常保持と停止を処理する / エラー発生条件（RESETで解除） / ①Stm A Axis001 絶対値位置決め エラー *)
Error_ST6_A_M[1] := (Stm_A_Rev_Axis000_MoveError OR Error_ST6_A_M[1]) AND NOT In_Sw_RESET;
(* Rung 30 *)
IF Error_ST6_A_M[1] THEN
    Retry[10] := TRUE;
    Out_TDC_Stop := TRUE;
END_IF;
(* Rung 31: #【A側ST7 排出異常】 / ワーク不一致・NG満杯・設定・回転異常 / RESETで解除、STARTで再確認 / Retry[11]：既存の停止・再試行経路 *)
Error_ST7_A_M[0] := (ST7_A_Dis2_M[11] OR ST7_A_Dis2_M[43] OR ST7_A_Dis2_M[44] OR Error_ST7_A_M[0]) AND NOT In_Sw_RESET;
(* Rung 32 *)
IF Error_ST7_A_M[0] THEN
    Retry[11] := TRUE;
    Out_TDC_Stop := TRUE;
END_IF;
(* Rung 33: 再試行：Retry[12] / 目的：原因別の異常保持と停止を処理する / エラー発生条件（RESETで解除） / ①軸異常 / ②非常停止状態（監視） / ③過負荷警告 *)
Error_ST7_A_M[1] := (RCON1_3_Error OR RCON1_5_Error OR Error_ST7_A_M[1]) AND NOT In_Sw_RESET;
(* Rung 34 *)
IF Error_ST7_A_M[1] THEN
    Retry[12] := TRUE;
    Out_TDC_Stop := TRUE;
END_IF;

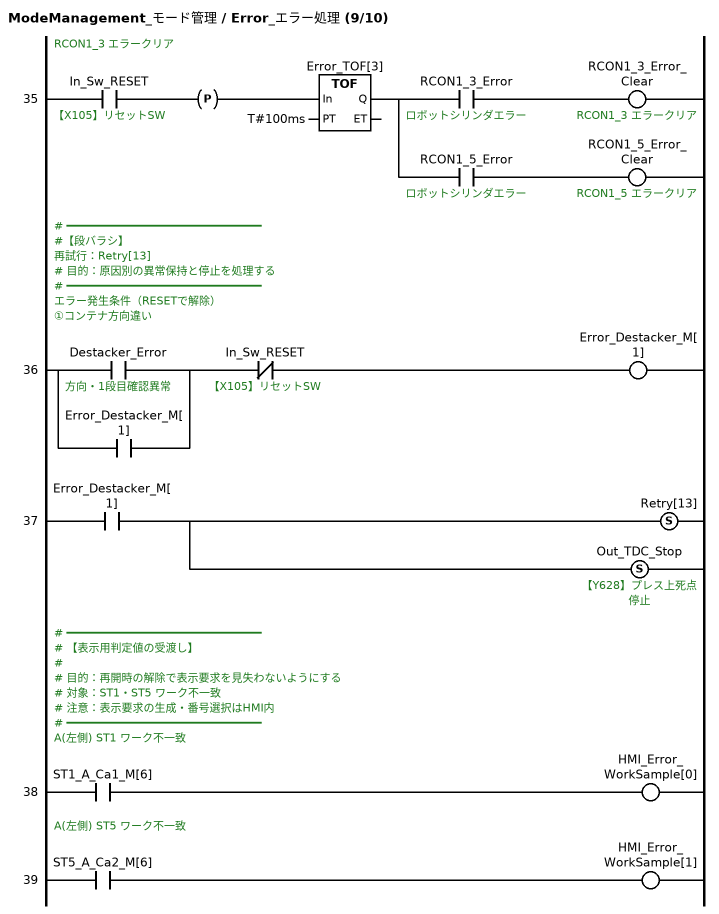
(* Rung 35: RCON1_3 エラークリア *)
_e47(CLK := In_Sw_RESET);
Error_TOF[3](In := _e47.Q, PT := T#100ms);
RCON1_3_Error_Clear := Error_TOF[3].Q AND RCON1_3_Error;
RCON1_5_Error_Clear := Error_TOF[3].Q AND RCON1_5_Error;
(* Rung 36: # ━━━━━━━━━━━━━━━━━━━━━━━━━━━━━━ / #【段バラシ】 / 再試行：Retry[13] / # 目的：原因別の異常保持と停止を処理する / # ━━━━━━━━━━━━━━━━━━━━━━━━━━━━━━ / エラー発生条件（RESETで解除） / ①コンテナ方向違い *)
Error_Destacker_M[1] := (Destacker_Error OR Error_Destacker_M[1]) AND NOT In_Sw_RESET;
(* Rung 37 *)
IF Error_Destacker_M[1] THEN
    Retry[13] := TRUE;
    Out_TDC_Stop := TRUE;
END_IF;
(* Rung 38: # ━━━━━━━━━━━━━━━━━━━━━━━━━━━━━━ / # 【表示用判定値の受渡し】 / # / # 目的：再開時の解除で表示要求を見失わないようにする / # 対象：ST1・ST5 ワーク不一致 / # 注意：表示要求の生成・番号選択はHMI内 / # ━━━━━━━━━━━━━━━━━━━━━━━━━━━━━━ / A(左側) ST1 ワーク不一致 *)
HMI_Error_WorkSample[0] := ST1_A_Ca1_M[6];
(* Rung 39: A(左側) ST5 ワーク不一致 *)
HMI_Error_WorkSample[1] := ST5_A_Ca2_M[6];

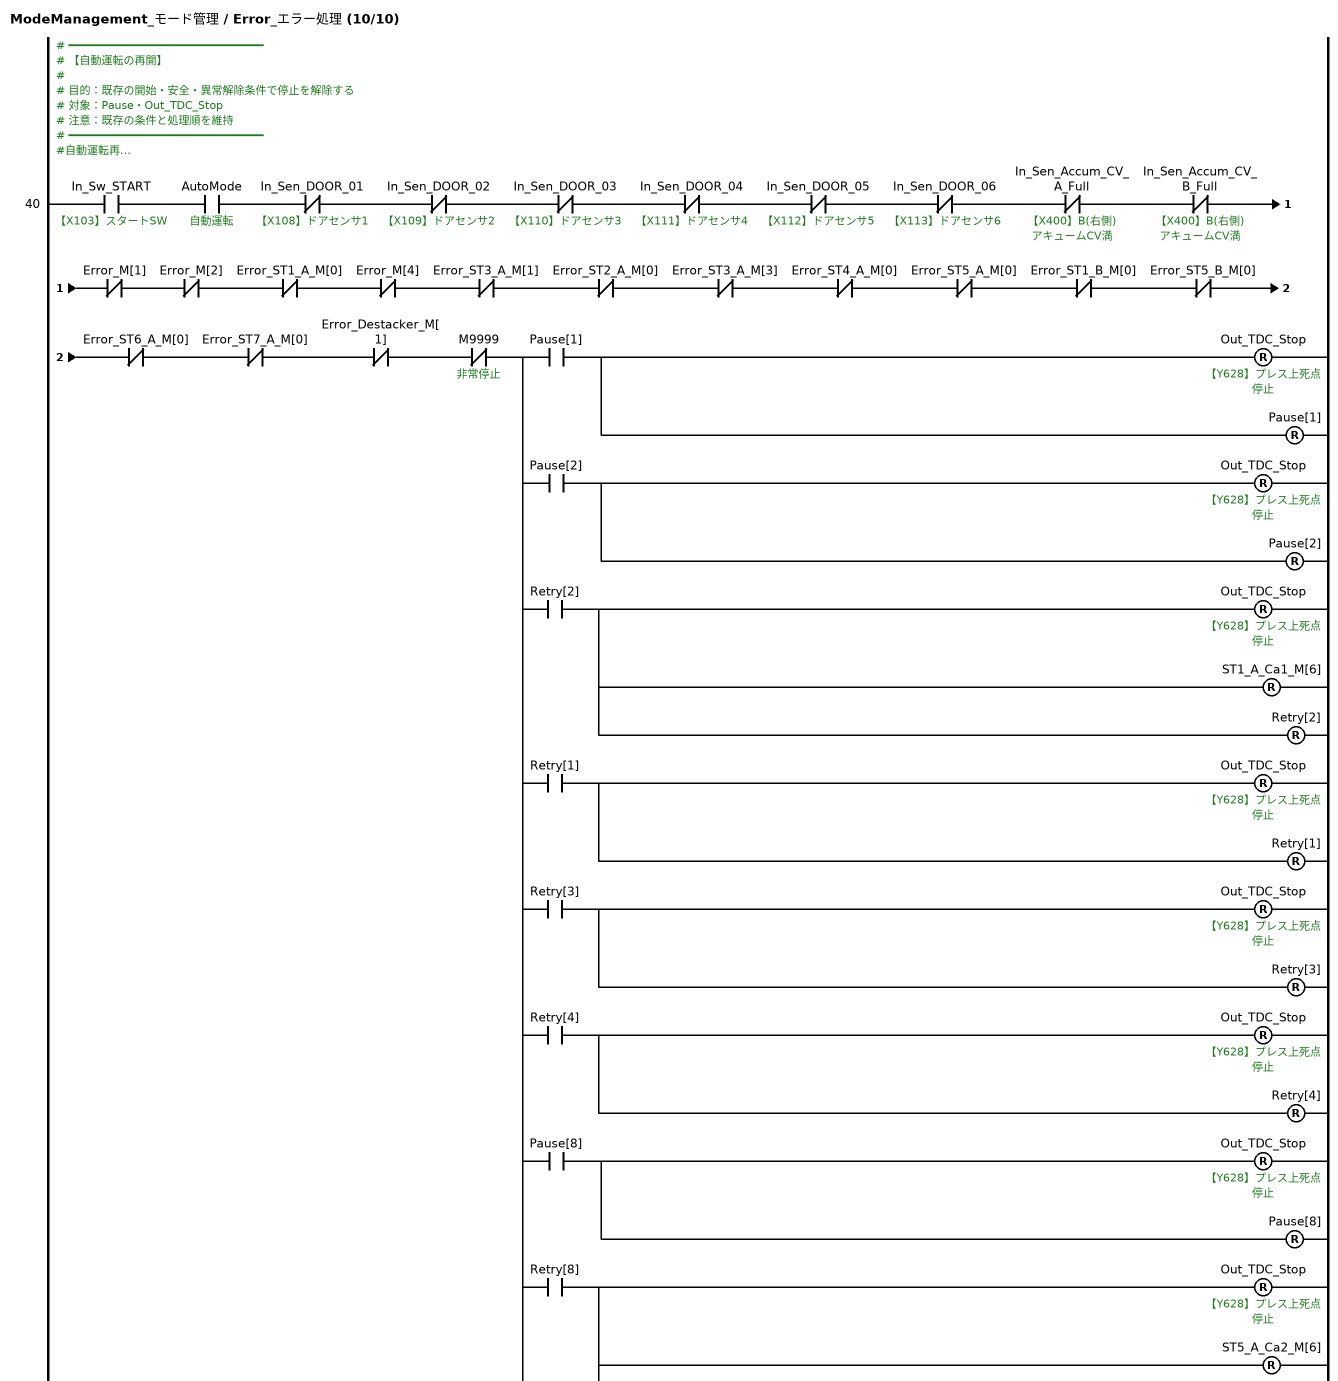

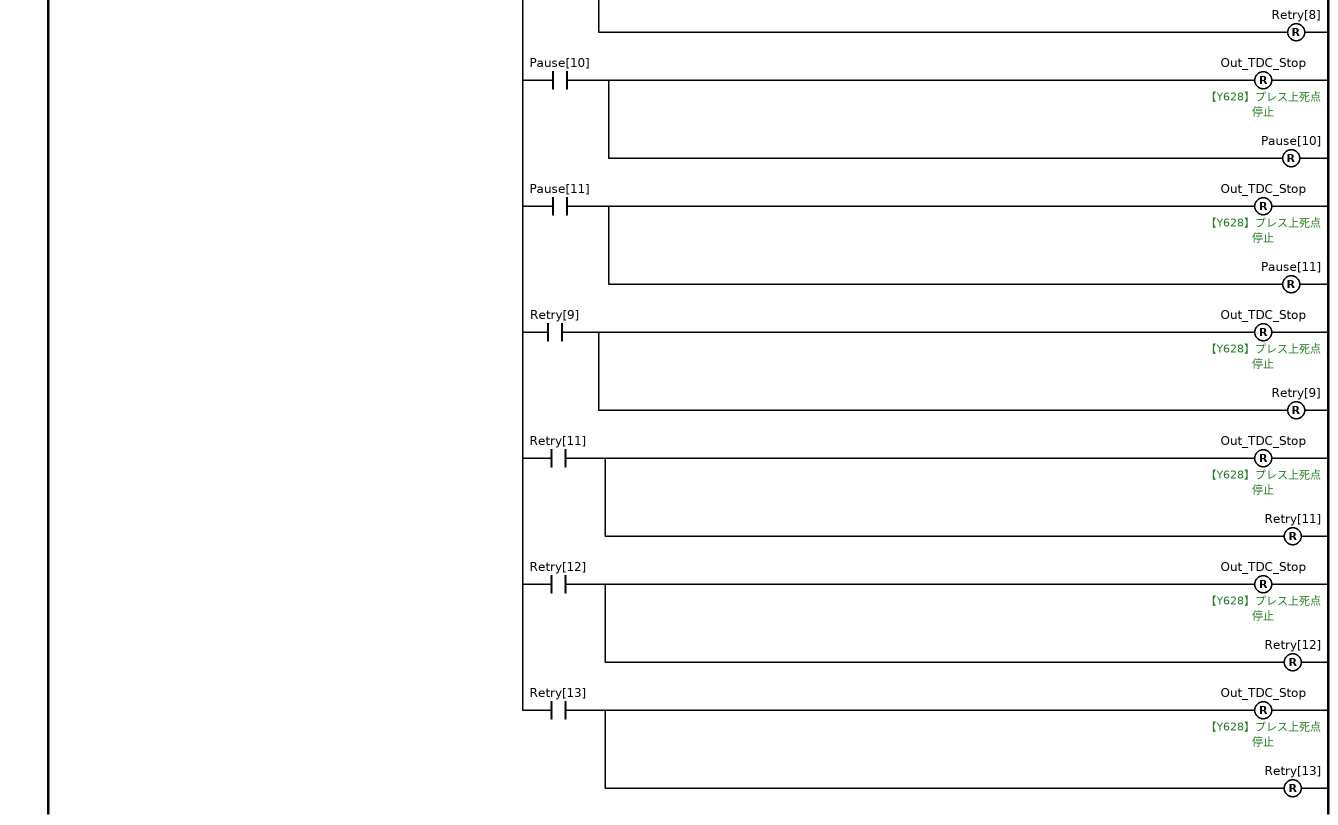
(* Rung 40: # ━━━━━━━━━━━━━━━━━━━━━━━━━━━━━━ / # 【自動運転の再開】 / # / # 目的：既存の開始・安全・異常解除条件で停止を解除する / # 対象：Pause・Out_TDC_Stop / # 注意：既存の条件と処理順を維持 / # ━━━━━━━━━━━━━━━━━━━━━━━━━━━━━━ / #自動運転再開 / 既存の開始・安全・異常・Pause解除条件を維持 *)
_p48 := In_Sw_START AND AutoMode AND NOT In_Sen_DOOR_01 AND NOT In_Sen_DOOR_02 AND NOT In_Sen_DOOR_03 AND NOT In_Sen_DOOR_04 AND NOT In_Sen_DOOR_05 AND NOT In_Sen_DOOR_06 AND NOT In_Sen_Accum_CV_A_Full AND NOT In_Sen_Accum_CV_B_Full AND NOT Error_M[1] AND NOT Error_M[2] AND NOT Error_ST1_A_M[0] AND NOT Error_M[4] AND NOT Error_ST3_A_M[1] AND NOT Error_ST2_A_M[0] AND NOT Error_ST3_A_M[3] AND NOT Error_ST4_A_M[0] AND NOT Error_ST5_A_M[0] AND NOT Error_ST1_B_M[0] AND NOT Error_ST5_B_M[0] AND NOT Error_ST6_A_M[0] AND NOT Error_ST7_A_M[0] AND NOT Error_Destacker_M[1] AND NOT M9999;
IF _p48 AND Pause[1] THEN
    Out_TDC_Stop := FALSE;
    Pause[1] := FALSE;
END_IF;
IF _p48 AND Pause[2] THEN
    Out_TDC_Stop := FALSE;
    Pause[2] := FALSE;
END_IF;
IF _p48 AND Retry[2] THEN
    Out_TDC_Stop := FALSE;
    ST1_A_Ca1_M[6] := FALSE;
    Retry[2] := FALSE;
END_IF;
IF _p48 AND Retry[1] THEN
    Out_TDC_Stop := FALSE;
    Retry[1] := FALSE;
END_IF;
IF _p48 AND Retry[3] THEN
    Out_TDC_Stop := FALSE;
    Retry[3] := FALSE;
END_IF;
IF _p48 AND Retry[4] THEN
    Out_TDC_Stop := FALSE;
    Retry[4] := FALSE;
END_IF;
IF _p48 AND Pause[8] THEN
    Out_TDC_Stop := FALSE;
    Pause[8] := FALSE;
END_IF;
IF _p48 AND Retry[8] THEN
    Out_TDC_Stop := FALSE;
    ST5_A_Ca2_M[6] := FALSE;
    Retry[8] := FALSE;
END_IF;
IF _p48 AND Pause[10] THEN
    Out_TDC_Stop := FALSE;
    Pause[10] := FALSE;
END_IF;
IF _p48 AND Pause[11] THEN
    Out_TDC_Stop := FALSE;
    Pause[11] := FALSE;
END_IF;
IF _p48 AND Retry[9] THEN
    Out_TDC_Stop := FALSE;
    Retry[9] := FALSE;
END_IF;
IF _p48 AND Retry[11] THEN
    Out_TDC_Stop := FALSE;
    Retry[11] := FALSE;
END_IF;
IF _p48 AND Retry[12] THEN
    Out_TDC_Stop := FALSE;
    Retry[12] := FALSE;
END_IF;
IF _p48 AND Retry[13] THEN
    Out_TDC_Stop := FALSE;
    Retry[13] := FALSE;
END_IF;
END_PROGRAM

PROGRAM Movements_動作
VAR
    Mo_M : BOOL;
    ST0_A_Sup_M : ARRAY[0..99] OF Bool;  (* [4] 原点位置移動完了 *)
    ST1_Ins_Cv_Rdy : BOOL;
    ST2_Ins_Cv_Rdy : BOOL;
    ST3_Ins_Cv_Rdy : BOOL;
    ST4_Ins_Cv_Rdy : BOOL;
    ST5_Ins_Cv_Rdy : BOOL;
    ST6_Ins_Cv_Rdy : BOOL;
    ST7_Ins_Cv_Rdy : BOOL;
    Ins_A_Cv_T : ARRAY[0..99] OF TON;
    ST1_A_Ca1_Rdy : BOOL;
    GT2_A_Inspection_GetTime : DATE_AND_TIME;
    GT2_A_Inspection_GetTime_ST : STRING[256];
    GT2_A_Inspection_GetTime_ST_Del : STRING[20];
    ST4_A_Rev1_Busy : BOOL;  (* ST4 A 動作中 *)
    ST6_A_Rev2_Busy : BOOL;  (* A(左側) ST6 反転2動作中 *)
    ST7_A_Dis2_Busy : BOOL;  (* ST7動作中 *)
    ST7_A_SF_M : ARRAY[0..99] OF Bool;  (* [2] フォルダ回転中; [1] フォルダ回転開始; [3] ターン戻要求; [4] ターン行要求; [5] 回転端位置正常 *)
    ST7_A_SF_Busy : BOOL;
    Destacker_TON : ARRAY[0..99] OF TON;
    BoxPacking_M : ARRAY[0..99] OF Bool;  (* 箱詰め工程; [1] 初回確認開始; [2] 初回確認完了; [3] 初回コンテナ状態判定; [4] 受渡位置・コンテナ到着; [5] コンテナ設置位置状態; [6] コンテナ排出位置状態; [7] コンテナ軸位置未確定; [8] Y1204 コンテナ排出戻; [9] コンテナ軸 初回設置移動; [10] コンテナ方向判定; [11] コンテナ方向OK; [12] 方向NGコンテナ 排出移動; [13] 初回コンテナ排出; [14] 初回コンテナ通過確認; [15] コンテナ軸 受渡位置移動; [16] 受渡位置・到着確認; [17] Y1206 箱入れチャック戻; [18] コンテナ軸 設置位置移動; [19] コンテナ設置完了; [20] 取出し先判定中; [21] A側取出し選択; [22] B側取出し選択; [23] 箱詰めZ 取出し準備上昇; [24] A側取出しXY移動; [25] A側取出しX完了; [26] A側取出しY完了; [27] A側取出しXY完了; [28] B側取出しXY移動; [29] B側取出しX完了; [30] B側取出しY完了; [31] B側取出しXY完了; [32] 箱詰めZ 取出し下降; [33] Y1207 取出しチャック行; [34] 箱詰めZ 取出し後上昇; [35] 箱内X位置選択・移動; [36] 箱内Y位置選択・移動; [37] 箱内X移動完了; [38] 箱内Y移動完了; [39] 箱内XY移動完了; [40] 箱詰めZ 箱内下降; [41] Y1206 箱内チャック戻; [42] 箱詰めZ 箱内配置後上昇; [43] コンテナ入数判定; [44] 80個未満・次取出し; [45] 80個・満杯排出; [46] コンテナ軸 満杯排出移動; [47] Y1205 満杯コンテナ排出行; [48] Y1204 満杯排出後戻; [49] コンテナ軸 排出後受渡戻 *)
    HMI_RCON2_2_OUT_TargetPos : ARRAY[0..99] OF LREAL;  (* RCON2_2 箱詰めX位置 [mm]; [1] A(左側)フォルダストック 取出しPos; [2] B(右側)フォルダストック 取出しPos; [3] 箱内X開始位置 [mm]：5個積みの1列目（設定値を入力） *)
    HMI_RCON2_5_OUT_TargetPos : ARRAY[0..99] OF LREAL;  (* RCON2_5 コンテナ軸位置 [mm]; [2] コンテナ設置Pos; [3] コンテナ排出Pos; [1] コンテナ受渡可能・セイフティ *)
    BoxPacking_Error : BOOL;  (* コンテナトレイ方向NG *)
    BoxPacking_TON : ARRAY[0..99] OF TON;
    A_SF_StackStepOffset : LREAL;  (* 積み段数－1 *)
    A_SF_StackDelta_mm : LREAL;  (* ピッチ×段数補正 [mm] *)
    A_SF_StackTarget_mm : LREAL;  (* 基準[3]＋積みピッチ補正 [mm] *)
    HMI_RCON2_3_OUT_TargetPos : ARRAY[0..99] OF LREAL;  (* RCON2_3 箱詰めY位置 [mm]; [1] A(左側)フォルダストック 取出しPos; [2] B(右側)フォルダストック 取出しPos; [3] 箱内Y開始位置 [mm]：4列×4行の1行目（設定値を入力） *)
    BoxPacking_A_Busy : BOOL;  (* A側取出し・箱内配置中 *)
    BoxPacking_B_Busy : BOOL;  (* B側 ストックフォルダ取出し中 *)
    BoxPacking_End : BOOL;  (* 満杯排出・軸戻り完了 *)
    BoxPacking_Init_Busy : BOOL;  (* 初回コンテナ確認中 *)
    BoxPacking_A_Pickup_Done : BOOL;  (* A側取出し・Z退避完了 *)
    Destacker_Init_Busy : BOOL;  (* 初回処理中 *)
    ST7_A_SF_Watch_TON : TON;  (* フォルダ回転10秒監視 *)
END_VAR
VAR_EXTERNAL
    ST0_Sup_Start : BOOL;  (* ST0_動作開始 *)
    M9999 : BOOL;
    Out_CYw_Sply_Pick_A_H_Auto : ARRAY[0..10] OF Bool;
    Out_CYw_Sply_Pick_A_H_Done : BOOL;
    Out_CYw_Sply_Slide_A_H_Auto : ARRAY[0..10] OF Bool;
    Out_CYw_Sply_Slide_A_H_Done : BOOL;
    Out_CYw_Sup_Chuck_A_Cl_H_Auto : ARRAY[0..10] OF Bool;
    Out_CYw_Sup_Chuck_A_Cl_H_Done : BOOL;
    In_Sen_Accum_CV_A_Arrival : BOOL;
    In_Sen_Work_A_Pos_00 : BOOL;
    Out_CYw_Sply_Pick_A_F_Auto : ARRAY[0..10] OF Bool;
    Out_CYw_Sply_Pick_A_F_Done : BOOL;
    Out_CYw_Sup_Chuck_A_Cl_F_Auto : ARRAY[0..10] OF Bool;
    Out_CYw_Sup_Chuck_A_Cl_F_Done : BOOL;
    Out_CYw_Sply_Slide_A_F_Auto : ARRAY[0..10] OF Bool;
    Out_CYw_Sply_Slide_A_F_Done : BOOL;
    Station_A_Data : ARRAY[0..8] OF sData;
    Cv_A_Data : ARRAY[0..8] OF sData;
    ST0_A_Sup_End : BOOL;  (* ST0 検査コンベア運転可 *)
    Out_CYS_Pos_01_Stopper_B_H_Auto : ARRAY[0..10] OF Bool;
    Out_CYS_Pos_02_Stopper_B_H_Auto : ARRAY[0..10] OF Bool;
    Out_CYS_Pos_03_Stopper_B_H_Auto : ARRAY[0..10] OF Bool;
    Out_CYS_Pos_04_Stopper_B_H_Auto : ARRAY[0..10] OF Bool;
    Out_CYS_Pos_05_Stopper_B_H_Auto : ARRAY[0..10] OF Bool;
    Out_CYS_Pos_06_Stopper_B_H_Auto : ARRAY[0..10] OF Bool;
    TimerQ_In_SenCY_Pos_01_Stopper_A_H : BOOL;
    TimerQ_In_SenCY_Pos_02_Stopper_A_H : BOOL;
    TimerQ_In_SenCY_Pos_03_Stopper_A_H : BOOL;
    TimerQ_In_SenCY_Pos_04_Stopper_A_H : BOOL;
    TimerQ_In_SenCY_Pos_05_Stopper_A_H : BOOL;
    TimerQ_In_SenCY_Pos_06_Stopper_A_H : BOOL;
    Out_Insp_Cv_A_Run_Auto : ARRAY[0..10] OF Bool;
    TimerQ_In_Sen_Work_A_Pos_01 : BOOL;
    TimerQ_In_Sen_Work_A_Pos_02 : BOOL;
    Pause : ARRAY[0..99] OF Bool;  (* [3] FH A(左側) ST1; [9] FH A(左側) ST5; [10] FH B(右側) ST1; [11] FH B(右側) ST5; [12] A(左側) ST6 反転2 ワーク不一致 *)
    TimerQ_In_Sen_Work_A_Pos_03 : BOOL;
    TimerQ_In_Sen_Work_A_Pos_04 : BOOL;
    TimerQ_In_Sen_Work_A_Pos_05 : BOOL;
    TimerQ_In_Sen_Work_A_Pos_06 : BOOL;
    TimerQ_In_Sen_Work_A_Pos_07 : BOOL;
    Out_CYS_Pos_01_Stopper_A_H_Auto : ARRAY[0..10] OF Bool;
    Out_CYS_Pos_02_Stopper_A_H_Auto : ARRAY[0..10] OF Bool;
    Out_CYS_Pos_03_Stopper_A_H_Auto : ARRAY[0..10] OF Bool;
    Out_CYS_Pos_04_Stopper_A_H_Auto : ARRAY[0..10] OF Bool;
    Out_CYS_Pos_05_Stopper_A_H_Auto : ARRAY[0..10] OF Bool;  (* [2] A(左側) ST5 カメラ2検査開始 *)
    Out_CYS_Pos_06_Stopper_A_H_Auto : ARRAY[0..10] OF Bool;  (* [1] A(左側)検査完了後; [2] A(左側) ST6 原点位置移動 *)
    Ins_A_Cv_M : ARRAY[0..99] OF Bool;
    Ins_A_Cv_Error : BOOL;  (* 検査コンベア ワーク不一致エラー *)
    TimerQ_In_Sen_Work_A_Pos_00 : BOOL;
    Out_CYS_Pos_01_Stopper_A_F_Auto : ARRAY[0..10] OF Bool;
    Out_CYS_Pos_02_Stopper_A_F_Auto : ARRAY[0..10] OF Bool;
    Out_CYS_Pos_03_Stopper_A_F_Auto : ARRAY[0..10] OF Bool;
    Out_CYS_Pos_04_Stopper_A_F_Auto : ARRAY[0..10] OF Bool;
    Out_CYS_Pos_05_Stopper_A_F_Auto : ARRAY[0..10] OF Bool;
    Out_CYS_Pos_06_Stopper_A_F_Auto : ARRAY[0..10] OF Bool;
    Ins_A_Next_Cycle : BOOL;  (* A(左側)検査コンベア 動作完了 *)
    ST0_A_Sup_Busy : BOOL;  (* ST0 稼働中 *)
    Ins_A_End : BOOL;  (* 検査完了 コンベア運転可能 *)
    Auto_A_Start : BOOL;
    Out_CYS_Pos_01_Stopper_A_H_Done : BOOL;
    FH_A_ST1_Auto : BOOL;
    FH_A_ST1_Done : BOOL;
    ST1_A_Ca1_Busy : BOOL;  (* ST1 A検査中 *)
    ST1_A_Ca1_End : BOOL;  (* ST1 A 動作完了 *)
    ST2_A_Hgt_Busy : BOOL;  (* ST2 A 動作中 *)
    Out_CYw_HgtInsp_Clp_A_H_Auto : ARRAY[0..10] OF Bool;
    Out_CYw_HgtInsp_Clp_A_H_Done : BOOL;
    Out_CYw_HgtInsp_Lf_A_H_Auto : ARRAY[0..10] OF Bool;
    Out_CYw_HgtInsp_Lf_A_H_Done : BOOL;
    Out_CYS_Pos_02_Stopper_A_H_Done : BOOL;
    Out_CYw_HgtInsp_Clp_A_F_Auto : ARRAY[0..10] OF Bool;
    Out_CYw_HgtInsp_Clp_A_F_Done : BOOL;
    Out_CYw_HgtInsp_Lf_A_F_Auto : ARRAY[0..10] OF Bool;
    Out_CYw_HgtInsp_Lf_A_F_Done : BOOL;
    DLEP1_GT2_A_Auto : BOOL;
    Hgt_A_ComputedValueData : LREAL;
    Hight_LowerLimit : LREAL;  (* 高さ検査 下限値 *)
    Hight_UpperLimit : LREAL;  (* 高さ検査 上限値 *)
    ST2_A_Hgt_End : BOOL;  (* 高さ検査完了 *)
    ST3_A_Dis1_Busy : BOOL;  (* ST3 A 動作中 *)
    Out_CYw_NG1_Srt_A_H_Auto : ARRAY[0..10] OF Bool;
    Out_CYw_NG1_Srt_A_H_Done : BOOL;
    Out_CYw_Rev_01_Pick_A_H_Auto : ARRAY[0..10] OF Bool;  (* 自動【Y710】A(左側)ST4 反転1ピックアップ戻： *)
    Out_CYw_Rev_01_Pick_A_H_Done : BOOL;  (* 【Y710】A(左側)ST4 反転1ピックアップ戻 動作完了 *)
    Out_CYw_NG1_Pick_A_H_Auto : ARRAY[0..10] OF Bool;
    Out_CYw_NG1_Pick_A_H_Done : BOOL;
    Out_CYw_NG1_Chk_A_H_Auto : ARRAY[0..10] OF Bool;
    Out_CYw_NG1_Chk_A_H_Done : BOOL;
    RCON1_1_Auto : ARRAY[0..99] OF Bool;  (* 自動移動要求; [1] 原点位置移動; [2] NG仕分け; [3] 動作完了後 原点位置移動 *)
    RCON1_1_OUT_TargetPos_mm : LREAL;  (* 目標位置 [mm] *)
    HMI_RCON1_1_OUT_TargetPos : ARRAY[0..99] OF LREAL;  (* HMI設定位置 [mm]; [1] 原点位置; [3] 高さNG位置; [4] カメラ キズNG位置; [5] カメラ 姿NG位置 *)
    RCON1_1_M : ARRAY[0..99] OF BOOL;  (* #A(左側) RCON1_1 NG1排出(上下); [1] 開始指令保持; [2] 予備 *)
    RCON1_1_MoveDone : BOOL;  (* 動作完了 *)
    Error_M : ARRAY[0..99] OF Bool;  (* [3] 未使用：Error_ST1_A_M[0]へ移行; [9] 未使用：Error_ST5_A_M[0]へ移行; [10] 未使用：Error_ST1_B_M[0]へ移行; [11] 未使用：Error_ST5_B_M[0]へ移行; [12] 未使用：Error_ST6_A_M[0]へ移行 *)
    ST1_A_Ca1_M : ARRAY[0..99] OF Bool;  (* [1] ST1 A カメラ1 検査開始; [2] 【Y720】A(左側) 位置1ストッパー 戻; [3] ワーク有無 判定; [4] ST1 A ワーク有; [5] ST1 A ワーク無; [6] A(左側) ST1 検査前ワーク不一致; [7] ST1 FH測定開始 *)
    ST2_A_Hgt_M : ARRAY[0..99] OF Bool;  (* [4] 【Y721】A(左側) 位置2ストッパー戻; [6] ST1 A ワーク有; [7] ST1 A ワーク無; [5] ワーク有無 判定; [9] 【Y703】A(左側) 高さ検査持上行; [10] 【Y701】A(左側) 高さ検査押え行; [11] A(左側) 高さ検査OK判定; [12] A(左側) 高さ検査NG判定; [2] 【Y701】A(左側) 高さ検査押え行; [8] ST3 検査前ワーク不一致エラー *)
    Out_CYS_Pos_03_Stopper_A_H_Done : BOOL;
    Out_CYw_NG1_Pick_A_F_Auto : ARRAY[0..10] OF Bool;
    Out_CYw_NG1_Pick_A_F_Done : BOOL;
    Out_CYw_NG1_Chk_A_F_Auto : ARRAY[0..10] OF Bool;
    Out_CYw_NG1_Chk_A_F_Done : BOOL;
    Out_CYw_NG1_Srt_A_F_Auto : ARRAY[0..10] OF Bool;
    Out_CYw_NG1_Srt_A_F_Done : BOOL;
    ST3_A_Dis1_End : BOOL;  (* 左NG1排出 完了 *)
    ST3_A_Dis1_M : ARRAY[0..99] OF Bool;  (* [7] 原点位置 移動開始; [6] 原点位置移動 データ転送; [5] 【Y722】A(左側) 位置3ストッパー戻; [4] 【Y706】A(左側) NG1チャック戻; [8] ワーク有無 / 検査前ワーク不一致 判定; [9] S3 A ワーク有 工程NG; [10] S3 A ワーク無  前工程OK; [14] 【Y704】A(左側) NG1ピックアップ戻 ; [24] 仕分け完了 *)
    ST4_A_Rev1_M : ARRAY[0..99] OF Bool;  (* [2] ワーク有無 / 検査前ワーク不一致 判定; [3] 【Y723】A(左側) 位置4ストッパー戻; [4] ST4 A ワーク有; [5] ST4 A ワーク無 / 前工程NG; [6] ST4 検査前ワーク不一致エラー; [10] A(左側) ST4 ワーク不一致エラー; [12] 【Y708】A(左側) ST4 反転1チャック閉 *)
    Stm_A_Rev_Axis000_MovePos_Degree : LREAL;
    HMI_Stm_A_Rev_Axis000_MovePos_Degree : ARRAY[0..99] OF LREAL;  (* A(左側)ステッピングモータ000 回転角度 *)
    Stm_A_Rev_Axis000_Auto : ARRAY[0..99] OF Bool;  (* [1] 原点位置移動 開始 *)
    Stm_A_Rev_Axis000_MoveAbsoluteDone : BOOL;
    Out_CYw_Rev_01_Pick_A_F_Auto : ARRAY[0..10] OF Bool;
    Out_CYw_Rev_01_Pick_A_F_Done : BOOL;
    Out_CYw_Disc_Chk_A_H_Auto : ARRAY[0..10] OF Bool;
    Out_CYw_Disc_Chk_A_H_Done : BOOL;
    Out_CYw_Rev_02_Chk_A_H_Auto : ARRAY[0..10] OF Bool;
    Out_CYw_Rev_02_Chk_A_H_Done : BOOL;
    Out_CYw_Rev_02_Chk_A_F_Auto : ARRAY[0..10] OF Bool;
    Out_CYw_Rev_01_Chk_A_F_Auto : ARRAY[0..10] OF Bool;
    Out_CYw_Rev_01_Chk_A_F_Done : BOOL;
    ST5_A_Ca2_M : ARRAY[0..99] OF Bool;  (* A(左側) ST5 カメラ2工程; [1] A(左側) ST5 カメラ2検査開始; [2] 【Y724】A(左側) ST5 ストッパー戻; [3] A(左側) ST5 ワーク有無判定; [4] A(左側) ST5 ワーク有; [5] A(左側) ST5 ワーク無; [6] A(左側) ST5 検査前ワーク不一致; [7] A(左側) ST5 FH測定開始 *)
    ST5_A_Ca2_Busy : BOOL;  (* A(左側) ST5 カメラ2検査中 *)
    ST5_A_Ca2_End : BOOL;  (* A(左側) ST5 カメラ2動作完了 *)
    FH_A_ST5_Auto : BOOL;  (* A(左側) ST5 FH自動測定 *)
    FH_A_ST5_Done : BOOL;  (* A(左側) ST5 画像検査完了 *)
    Out_CYS_Pos_05_Stopper_A_H_Done : BOOL;  (* 【Y724】A(左側) 位置5ストッパー戻 動作完了 *)
    Out_CYw_Rev_01_Chk_A_H_Auto : ARRAY[0..10] OF Bool;  (* 自動【Y708】A(左側)ST4 反転1チャック閉： *)
    Out_CYw_Rev_01_Chk_A_H_Done : BOOL;  (* 【Y708】A(左側)ST4 反転1チャック閉 動作完了 *)
    HMI_Stm_A_Rev_Axis001_MovePos_Degree : ARRAY[0..99] OF LREAL;  (* A(左側) ST6 反転2設定角度; [1] A(左側) ST6 原点位置設定角度; [2] A(左側) ST6 反転位置設定角度 *)
    Out_CYw_Rev_02_Chk_A_F_Done : BOOL;  (* 【Y713】A(左側)ST6 反転2チャック開 行 動作完了 *)
    Out_CYw_Rev_02_Pick_A_F_Auto : ARRAY[0..10] OF Bool;  (* 自動【Y715】A(左側)ST6 反転2ピックアップ行 ：; [1] A(左側) ST6 反転前行; [2] A(左側) ST6 設置行 *)
    Out_CYw_Rev_02_Pick_A_F_Done : BOOL;  (* 【Y715】A(左側)ST6 反転2ピックアップ行 動作完了 *)
    Out_CYw_Rev_02_Pick_A_H_Auto : ARRAY[0..10] OF Bool;  (* 自動【Y714】A(左側)ST6 反転2ピックアップ戻 ：; [1] A(左側) ST6 反転前戻; [2] A(左側) ST6 設置後戻 *)
    Out_CYw_Rev_02_Pick_A_H_Done : BOOL;  (* 【Y714】A(左側)ST6 反転2ピックアップ戻 動作完了 *)
    Stm_A_Rev_Axis001_Auto : ARRAY[0..99] OF Bool;  (* A(左側) ST6 反転2自動指令; [1] A(左側) ST6 原点位置移動開始 *)
    Stm_A_Rev_Axis001_MoveAbsoluteDone : BOOL;  (* A(左側) ST6 反転2位置決め完了 *)
    Stm_A_Rev_Axis001_MovePos_Degree : LREAL;  (* A(左側) ST6 反転2指令角度 *)
    ST6_A_Rev2_M : ARRAY[0..99] OF Bool;
    RCON1_5_Auto : ARRAY[0..99] OF Bool;  (* 自動移動要求; [1] 初期安全上昇; [2] コンベア回収下降; [3] 保持後安全上昇; [4] 仕分け先へ下降; [5] 解放後安全上昇 *)
    HMI_RCON1_5_OUT_TargetPos : ARRAY[0..99] OF LREAL;  (* RCON1_5 目標位置 [mm]：; [1] 安全上昇位置; [2] コンベア回収下降位置; [3] OK積み1段目の基準; [4] 旧段別位置4：現在未使用; [5] 旧段別位置5：現在未使用; [6] 旧段別位置6：現在未使用; [7] キズNG下降位置; [8] 姿NG下降位置 *)
    RCON1_5_MoveDone : BOOL;
    Out_CYw_Ejc_Hldr_Feed_A_H_Auto : ARRAY[0..10] OF Bool;
    Out_CYw_Ejc_Hldr_Feed_A_H_Done : BOOL;
    HMI_RCON1_3_OUT_TargetPos : ARRAY[0..99] OF LREAL;  (* RCON1_3 SF/NG2仕分け(左右) 目標位置 [mm]： *)
    RCON1_3_Auto : ARRAY[0..99] OF Bool;
    RCON1_3_MoveDone : BOOL;
    ST7_A_Dis2_M : ARRAY[0..99] OF Bool;  (* [9] ワーク有; [10] ワーク無; [11] 有無・NG満杯異常; [12] 回収下降位置転送; [13] 回収下降要求; [14] ワーク保持; [15] 保持後上昇位置転送; [16] 保持後上昇要求; [17] 仕分け位置選択; [18] OK選択; [19] キズNG選択; [20] 姿NG選択; [21] OK送り行開始; [22] 仕分け左右移動中; [23] 下降位置選択; [24] OK積み位置; [25] キズNG下降位置; [26] 姿NG下降位置; [27] 配置下降要求; [28] ワーク解放; [29] 解放後上昇位置転送; [30] 解放後上昇要求; [31] 左右原点位置転送; [32] 左右原点移動要求; [33] 最後の送り戻; [1] 排出動作開始; [2] 初期チャック戻; [3] 初期上昇位置転送; [4] 初期上昇要求; [5] 初期左右位置転送; [6] 初期左右移動要求; [7] 初期送り戻; [8] ワーク有無判定; [42] 今回ワーク加算済み; [43] 積み設定・判定異常; [44] フォルダ回転異常; [45] ワーク回収開始許可; [46] 今回の初期位置確認済み; [34] 初期上昇 前完了解除; [35] 初期左右 前完了解除; [36] 回収下降 前完了解除; [37] 保持後上昇 前完了解除; [38] 仕分け左右 前完了解除; [39] 配置下降 前完了解除; [40] 解放後上昇 前完了解除; [41] 左右戻り 前完了解除 *)
    RCON1_3_OUT_TargetPos_mm : LREAL;
    A_SF_CT : INT;  (* A(左側) ストックフォルダカウント *)
    TimerQ_In_Sen_SH_B_Ent : BOOL;
    TimerQ_In_Sen_SH_B_Ext : BOOL;
    RCON1_5_ActualPos_mm : LREAL;
    RCON1_5_SafePos_mm : LREAL;
    Out_CYw_SH_A_Turn_F_Auto : ARRAY[0..10] OF Bool;
    TimerQ_In_SenCY_SH_A_Turn_F : BOOL;
    Out_CYw_SH_A_Turn_H_Auto : ARRAY[0..10] OF Bool;
    TimerQ_In_SenCY_SH_A_Turn_H : BOOL;
    Out_CYw_SH_A_Turn_H_Done : BOOL;
    Out_CYw_SH_A_Turn_F_Done : BOOL;
    Out_CYw_Ejc_Hldr_Feed_A_F_Auto : ARRAY[0..10] OF Bool;
    Out_CYw_Ejc_Hldr_Feed_A_F_Done : BOOL;
    Out_CYw_Disc_Chk_A_F_Auto : ARRAY[0..10] OF Bool;
    Out_CYw_Disc_Chk_A_F_Done : BOOL;
    RCON1_5_OUT_TargetPos_mm : LREAL;
    ST7_A_Dis2_End : BOOL;  (* ST7 A 動作完了 *)
    In_Sen_NG2_Tray_B_Full : BOOL;
    TimerQ_In_Sen_NG2_Tray_B_Full : BOOL;
    TimerQ_In_Sen_NG1_Tray_B_Full : BOOL;
    ST7_A_SF_Wait_Pickup : BOOL;  (* フォルダストック取出し待ち *)
    Error_ST7_A_Source_M : ARRAY[0..4] OF BOOL;  (* #A(左側) ST7 発生理由（内部保持）; [3] ワーク不一致; [4] 満杯（既存B側入力） *)
    Retry : ARRAY[0..99] OF BOOL;
    TimerQ_In_Sen_NG2_Tray_A_Full : BOOL;
    ST6_A_Rev2_End : BOOL;  (* A(左側) ST6 反転2動作完了 *)
    ST4_A_Rev_End : BOOL;
    Auto_Com_Start : BOOL;
    Destacker_M : ARRAY[0..99] OF Bool;  (* 段バラシ工程; [26] 初回確認済み; [27] 初回安全 前完了解除; [28] 初回1段 前完了解除; [29] 初回戻り 前完了解除; [30] 1段目 前完了解除; [31] 2段目 前完了解除; [32] 排出 前完了解除; [1] 初回確認開始; [2] 初回の爪保持; [3] 初回の位置判定; [4] 初回安全位置あり; [5] 初回安全位置なし; [6] 初回の爪戻し; [7] 初回安全位置移動; [8] 初回1段目移動; [9] 初回コンテナ保持; [10] 初回安全位置戻り; [11] 初回の送り戻し; [12] 通常サイクル開始; [13] 送り戻り待ち; [14] コンテナ確認中; [15] コンテナ確認OK; [16] 1段目位置へ移動; [17] コンテナ切り離し; [18] 段積み判定; [19] 2段以上; [20] 1段のみ; [21] 2段目位置へ移動; [22] 上段コンテナ保持; [23] 安全・排出位置移動; [24] 送り行待ち; [25] 送り戻り待ち *)
    Out_CYw_Sep_Claw_F_Auto : ARRAY[0..10] OF Bool;
    Out_CYw_Sep_Claw_F_Done : BOOL;
    RCON2_1_OUT_TargetPos_mm : LREAL;
    HMI_RCON2_1_OUT_TargetPos : ARRAY[0..99] OF LREAL;  (* 段バラシ 目標位置 [mm] *)
    RCON2_1_Auto : ARRAY[0..99] OF Bool;
    TimerQ_In_Sen_Supply_Container_Exist : BOOL;
    TimerQ_In_SenCY_Empty_Container_CY_H : BOOL;
    TimerQ_In_Sen_Destacker_Stage_01_Exist : BOOL;
    TimerQ_In_Sen_Destacker_Stage_02_Exist : BOOL;
    BoxPacking_Busy : BOOL;  (* 箱詰め動作中 *)
    RCON2_1_MoveDone : BOOL;
    TimerQ_In_Sen_Container_Direction_Check : BOOL;
    Out_CYw_Sep_Claw_H_Auto : ARRAY[0..10] OF Bool;
    Out_CYw_Sep_Claw_H_Done : BOOL;
    Destacker_End : BOOL;  (* 1サイクル完了 *)
    RCON2_1_ActualPos_mm : LREAL;
    Out_CYw_Ejc_Cont_F_Auto : ARRAY[0..10] OF Bool;
    Out_CYw_Ejc_Cont_F_Done : BOOL;
    Out_CYw_Ejc_Cont_H_Auto : ARRAY[0..10] OF Bool;
    Out_CYw_Empty_Container_CY_H_Auto : ARRAY[0..10] OF Bool;
    Out_CYw_Empty_Container_CY_H_Done : BOOL;
    TimerQ_In_SenCY_Empty_Container_CY_F : BOOL;
    Out_CYw_Empty_Container_CY_F_Auto : ARRAY[0..10] OF Bool;
    RCON2_2_ActualPos_mm : LREAL;
    RCON2_5_ActualPos_mm : LREAL;
    Out_CYw_Empty_Container_CY_F_Done : BOOL;
    In_Sen_Container_Arrival : BOOL;
    TimerQ_In_Sen_Container_Arrival : BOOL;
    Destacker_Error : BOOL;  (* 方向・1段目確認異常 *)
    RCON2_5_OUT_TargetPos_mm : LREAL;
    RCON2_5_Auto : ARRAY[0..99] OF Bool;
    RCON2_5_MoveDone : BOOL;
    TimerQ_In_Sen_Tray_Direction_Check : BOOL;
    Out_CYw_Ejc_Cont_H_Done : BOOL;
    TimerQ_In_Sen_Container_Pass : BOOL;
    ST7_B_SF_Wait_Pickup : BOOL;  (* フォルダストックB取出し待ち *)
    RCON2_4_OUT_TargetPos_mm : LREAL;
    RCON2_4_Auto : ARRAY[0..99] OF Bool;
    HMI_A_SF_StackPitch_mm : LREAL;  (* 左SF積みピッチ [mm] *)
    A_Total_CT : INT;  (* A(左側)生産数 *)
    HMI_RCON2_4_OUT_TargetPos : ARRAY[0..99] OF LREAL;  (* RCON2_4 箱詰めZ位置 [mm]; [1] セイフティPos *)
    RCON2_2_OUT_TargetPos_mm : LREAL;
    RCON2_3_OUT_TargetPos_mm : LREAL;
    RCON2_2_Auto : ARRAY[0..99] OF Bool;
    RCON2_3_Auto : ARRAY[0..99] OF Bool;
    RCON2_2_MoveDone : BOOL;
    RCON2_3_MoveDone : BOOL;
    Out_CYw_Box_Chuck_F_Auto : ARRAY[0..10] OF Bool;
    Out_CYw_Box_Chuck_F_Done : BOOL;
    Out_CYw_Box_Chuck_H_Auto : ARRAY[0..10] OF Bool;
    Out_CYw_Box_Chuck_H_Done : BOOL;
    Box_Total_CT : INT;  (* コンテナ入数 *)
    HMI_Box_X_Pitch_mm : LREAL;  (* 箱詰めX方向の1ピッチ [mm]：符号付き。正=座標増、負=座標減。使用前に設定。 *)
    HMI_Box_Y_Pitch_mm : LREAL;  (* 箱詰めY方向の1ピッチ [mm]：符号付き。正=座標増、負=座標減。使用前に設定。 *)
    RCON2_4_MoveDone : BOOL;
    TimerQ_In_Sen_SH_A_Ent : BOOL;  (* 【X214】：A側積み側5個有 *)
    TimerQ_In_Sen_SH_A_Ext : BOOL;  (* 【X215】：A側取出し側5個有 *)
    In_Sw_RESET : BOOL;  (* リセットSW *)
END_VAR
VAR
    _e1 : R_TRIG;
    _p2 : BOOL;
    _e3 : R_TRIG;
    _e4 : R_TRIG;
    _p5 : BOOL;
    _e6 : R_TRIG;
    _e7 : R_TRIG;
    _p8 : BOOL;
    _p9 : BOOL;
    _p10 : BOOL;
    _p11 : BOOL;
    _p12 : BOOL;
    _p13 : BOOL;
    _p14 : BOOL;
    _p15 : BOOL;
    _e16 : R_TRIG;
    _p17 : BOOL;
    _p18 : BOOL;
    _p19 : BOOL;
    _p20 : BOOL;
    _p21 : BOOL;
    _p22 : BOOL;
    _p23 : BOOL;
    _p24 : BOOL;
    _p25 : BOOL;
    _p26 : BOOL;
    _p27 : BOOL;
    _p28 : BOOL;
    _e29 : R_TRIG;
    _p30 : BOOL;
    _e31 : R_TRIG;
    _p32 : BOOL;
    _p33 : BOOL;
    _p34 : BOOL;
    _p35 : BOOL;
    _p36 : BOOL;
    _e37 : R_TRIG;
    _p38 : BOOL;
    _p39 : BOOL;
    _p40 : BOOL;
    _p41 : BOOL;
    _e42 : R_TRIG;
    _p43 : BOOL;
    _p44 : BOOL;
    _p45 : BOOL;
    _p46 : BOOL;
    _p47 : BOOL;
    _e48 : R_TRIG;
    _p49 : BOOL;
    _p50 : BOOL;
    _p51 : BOOL;
    _p52 : BOOL;
    _p53 : BOOL;
    _p54 : BOOL;
    _p55 : BOOL;
    _p56 : BOOL;
    _p57 : BOOL;
    _p58 : BOOL;
    _p59 : BOOL;
    _e60 : R_TRIG;
    _p61 : BOOL;
    _p62 : BOOL;
    _p63 : BOOL;
    _e64 : R_TRIG;
    _p65 : BOOL;
    _p66 : BOOL;
    _p67 : BOOL;
    _p68 : BOOL;
    _p69 : BOOL;
    _p70 : BOOL;
    _p71 : BOOL;
    _p72 : BOOL;
    _p73 : BOOL;
    _e74 : R_TRIG;
    _p75 : BOOL;
    _p76 : BOOL;
    _e77 : R_TRIG;
    _p78 : BOOL;
    _p79 : BOOL;
    _p80 : BOOL;
    _e81 : R_TRIG;
    _p82 : BOOL;
    _p83 : BOOL;
    _p84 : BOOL;
    _p85 : BOOL;
    _p86 : BOOL;
    _p87 : BOOL;
    _p88 : BOOL;
    _p89 : BOOL;
    _e90 : R_TRIG;
    _p91 : BOOL;
    _p92 : BOOL;
    _p93 : BOOL;
    _p94 : BOOL;
    _e95 : R_TRIG;
    _p96 : BOOL;
    _p97 : BOOL;
    _p98 : BOOL;
    _p99 : BOOL;
    _p100 : BOOL;
    _p101 : BOOL;
    _p102 : BOOL;
    _p103 : BOOL;
    _p104 : BOOL;
    _p105 : BOOL;
    _p106 : BOOL;
    _p107 : BOOL;
    _e108 : R_TRIG;
    _p109 : BOOL;
    _p110 : BOOL;
    _p111 : BOOL;
    _e112 : R_TRIG;
    _p113 : BOOL;
    _p114 : BOOL;
    _p115 : BOOL;
    _e116 : R_TRIG;
    _p117 : BOOL;
    _p118 : BOOL;
    _p119 : BOOL;
    _p120 : BOOL;
    _p121 : BOOL;
    _p122 : BOOL;
    _p123 : BOOL;
    _p124 : BOOL;
    _p125 : BOOL;
    _p126 : BOOL;
    _e127 : R_TRIG;
    _p128 : BOOL;
    _p129 : BOOL;
    _p130 : BOOL;
    _p131 : BOOL;
    _p132 : BOOL;
    _p133 : BOOL;
    _p134 : BOOL;
    _p135 : BOOL;
    _p136 : BOOL;
    _p137 : BOOL;
    _p138 : BOOL;
    _p139 : BOOL;
    _p140 : BOOL;
    _p141 : BOOL;
    _p142 : BOOL;
    _p143 : BOOL;
    _p144 : BOOL;
    _p145 : BOOL;
    _p146 : BOOL;
    _p147 : BOOL;
    _p148 : BOOL;
    _p149 : BOOL;
    _e150 : R_TRIG;
    _p151 : BOOL;
    _e152 : R_TRIG;
    _p153 : BOOL;
    _p154 : BOOL;
    _p155 : BOOL;
    _p156 : BOOL;
    _p157 : BOOL;
    _p158 : BOOL;
    _p159 : BOOL;
    _p160 : BOOL;
    _p161 : BOOL;
    _p162 : BOOL;
    _p163 : BOOL;
    _p164 : BOOL;
    _p165 : BOOL;
    _p166 : BOOL;
    _p167 : BOOL;
    _p168 : BOOL;
    _p169 : BOOL;
    _e170 : R_TRIG;
END_VAR

(* Section Ins_A_Cv_左検査Cv: ladder, written here as Structured Text *)

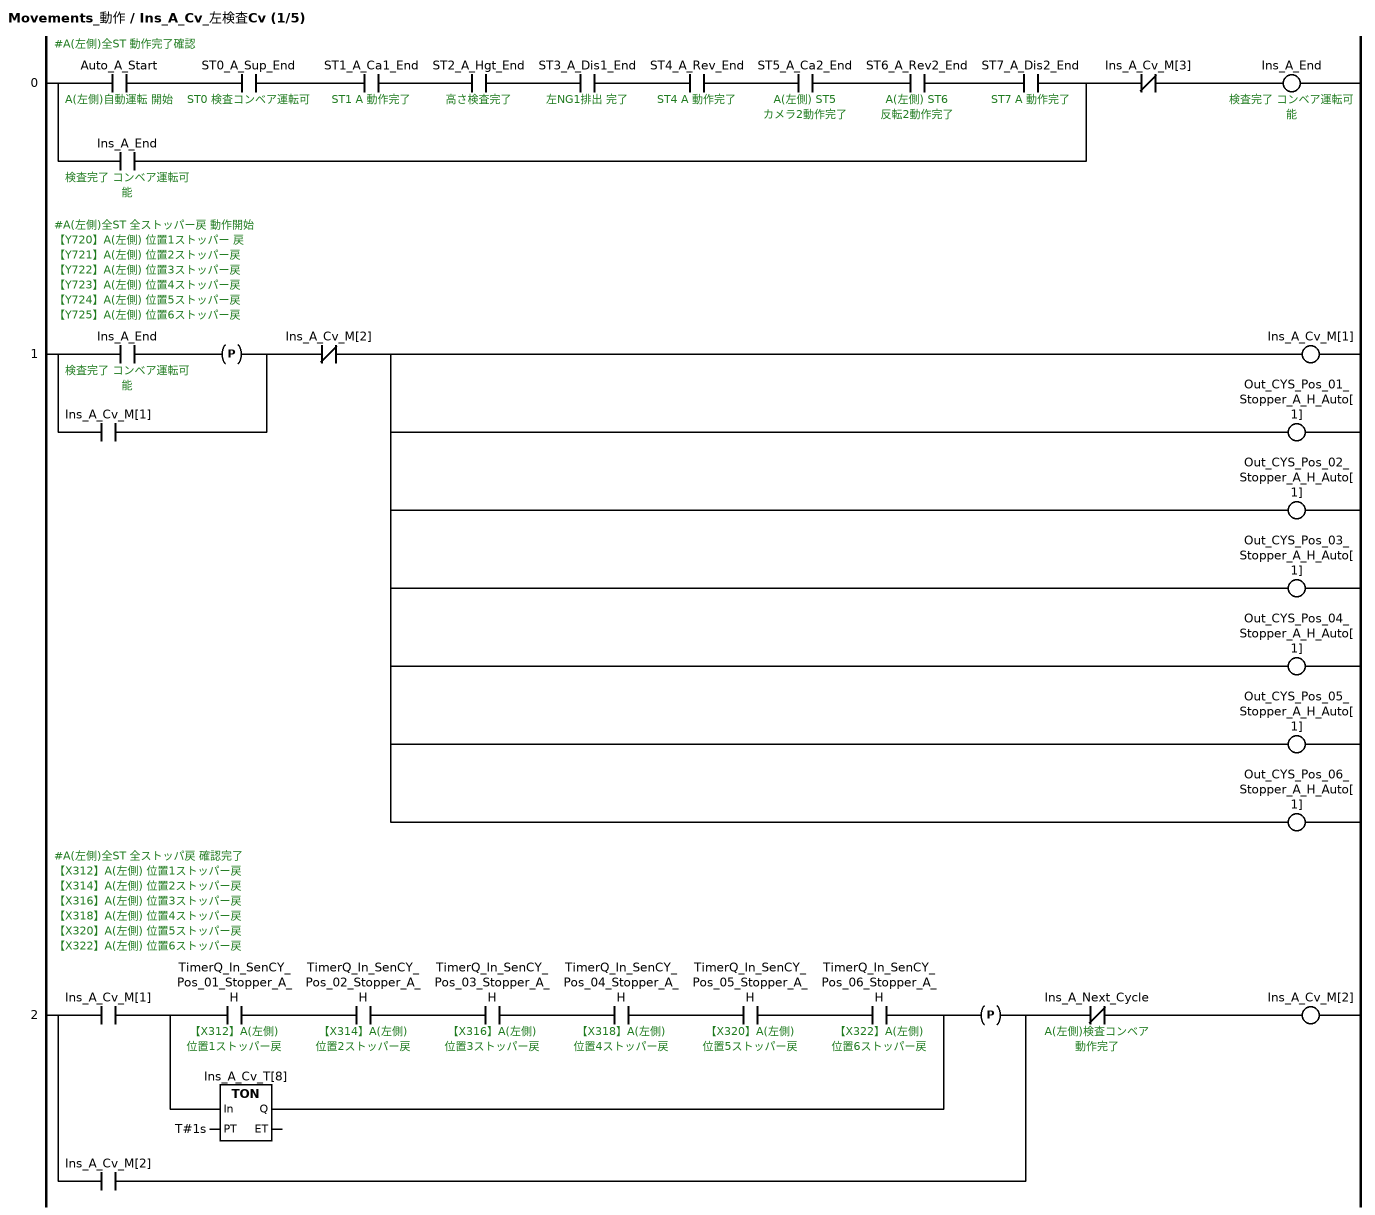
(* Rung 0: #A(左側)全ST 動作完了確認 *)
Ins_A_End := ((Auto_A_Start AND ST0_A_Sup_End AND ST1_A_Ca1_End AND ST2_A_Hgt_End AND ST3_A_Dis1_End AND ST4_A_Rev_End AND ST5_A_Ca2_End AND ST6_A_Rev2_End AND ST7_A_Dis2_End) OR Ins_A_End) AND NOT Ins_A_Cv_M[3];
(* Rung 1: #A(左側)全ST 全ストッパー戻 動作開始 / 【Y720】A(左側) 位置1ストッパー 戻 / 【Y721】A(左側) 位置2ストッパー戻 / 【Y722】A(左側) 位置3ストッパー戻 / 【Y723】A(左側) 位置4ストッパー戻 / 【Y724】A(左側) 位置5ストッパー戻 / 【Y725】A(左側) 位置6ストッパー戻 *)
_e1(CLK := Ins_A_End);
_p2 := (_e1.Q OR Ins_A_Cv_M[1]) AND NOT Ins_A_Cv_M[2];
Ins_A_Cv_M[1] := _p2;
Out_CYS_Pos_01_Stopper_A_H_Auto[1] := _p2;
Out_CYS_Pos_02_Stopper_A_H_Auto[1] := _p2;
Out_CYS_Pos_03_Stopper_A_H_Auto[1] := _p2;
Out_CYS_Pos_04_Stopper_A_H_Auto[1] := _p2;
Out_CYS_Pos_05_Stopper_A_H_Auto[1] := _p2;
Out_CYS_Pos_06_Stopper_A_H_Auto[1] := _p2;
(* Rung 2: #A(左側)全ST 全ストッパ戻 確認完了 / 【X312】A(左側) 位置1ストッパー戻 / 【X314】A(左側) 位置2ストッパー戻 / 【X316】A(左側) 位置3ストッパー戻 / 【X318】A(左側) 位置4ストッパー戻 / 【X320】A(左側) 位置5ストッパー戻 / 【X322】A(左側) 位置6ストッパー戻 *)
Ins_A_Cv_T[8](In := Ins_A_Cv_M[1], PT := T#1s);
_e3(CLK := (Ins_A_Cv_M[1] AND TimerQ_In_SenCY_Pos_01_Stopper_A_H AND TimerQ_In_SenCY_Pos_02_Stopper_A_H AND TimerQ_In_SenCY_Pos_03_Stopper_A_H AND TimerQ_In_SenCY_Pos_04_Stopper_A_H AND TimerQ_In_SenCY_Pos_05_Stopper_A_H AND TimerQ_In_SenCY_Pos_06_Stopper_A_H) OR Ins_A_Cv_T[8].Q);
Ins_A_Cv_M[2] := (_e3.Q OR Ins_A_Cv_M[2]) AND NOT Ins_A_Next_Cycle;

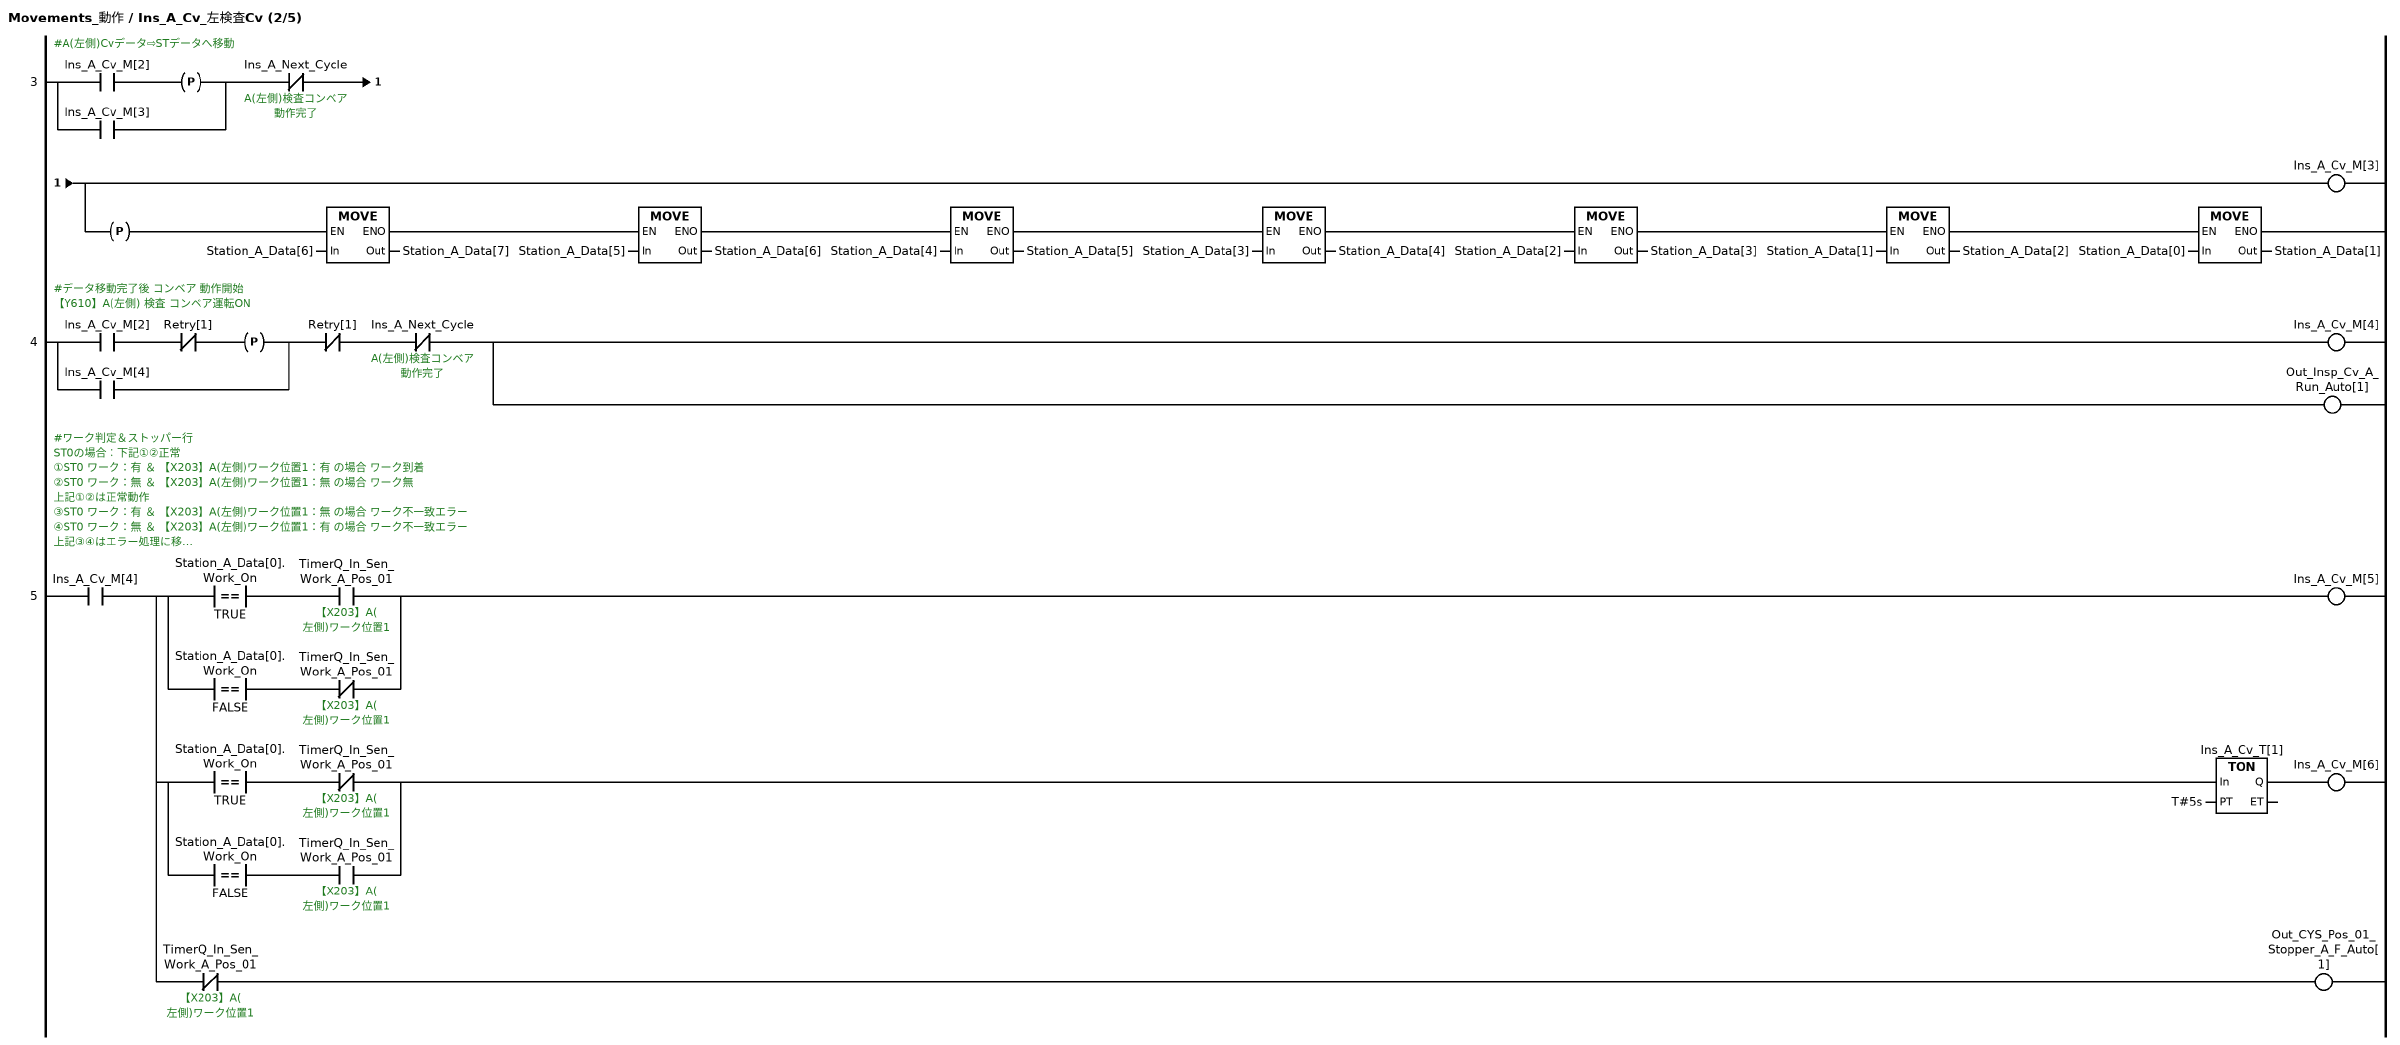
(* Rung 3: #A(左側)Cvデータ⇨STデータへ移動 *)
_e4(CLK := Ins_A_Cv_M[2]);
_p5 := (_e4.Q OR Ins_A_Cv_M[3]) AND NOT Ins_A_Next_Cycle;
Ins_A_Cv_M[3] := _p5;
_e6(CLK := _p5);
IF _e6.Q THEN
    Station_A_Data[7] := Station_A_Data[6];
    Station_A_Data[6] := Station_A_Data[5];
    Station_A_Data[5] := Station_A_Data[4];
    Station_A_Data[4] := Station_A_Data[3];
    Station_A_Data[3] := Station_A_Data[2];
    Station_A_Data[2] := Station_A_Data[1];
    Station_A_Data[1] := Station_A_Data[0];
END_IF;
(* Rung 4: #データ移動完了後 コンベア 動作開始 / 【Y610】A(左側) 検査 コンベア運転ON *)
_e7(CLK := Ins_A_Cv_M[2] AND NOT Retry[1]);
_p8 := (_e7.Q OR Ins_A_Cv_M[4]) AND NOT Retry[1] AND NOT Ins_A_Next_Cycle;
Ins_A_Cv_M[4] := _p8;
Out_Insp_Cv_A_Run_Auto[1] := _p8;
(* Rung 5: #ワーク判定＆ストッパー行 / ST0の場合：下記①②正常 / ①ST0 ワーク：有 ＆ 【X203】A(左側)ワーク位置1：有 の場合 ワーク到着 / ②ST0 ワーク：無 ＆ 【X203】A(左側)ワーク位置1：無 の場合 ワーク無 / 上記①②は正常動作 / ③ST0 ワーク：有 ＆ 【X203】A(左側)ワーク位置1：無 の場合 ワーク不一致エラー / ④ST0 ワーク：無 ＆ 【X203】A(左側)ワーク位置1：有 の場合 ワーク不一致エラー / 上記③④はエラー処理に移動 / ⑤【X203】A(左側)ワーク位置1：無 の場合 / 【Y720】A(左側) 位置1ストッパー 行 *)
_p9 := Ins_A_Cv_M[4];
Ins_A_Cv_M[5] := Ins_A_Cv_M[4] AND (((Station_A_Data[0].Work_On = TRUE) AND TimerQ_In_Sen_Work_A_Pos_01) OR ((Station_A_Data[0].Work_On = FALSE) AND NOT TimerQ_In_Sen_Work_A_Pos_01));
Ins_A_Cv_T[1](In := _p9 AND (((Station_A_Data[0].Work_On = TRUE) AND NOT TimerQ_In_Sen_Work_A_Pos_01) OR ((Station_A_Data[0].Work_On = FALSE) AND TimerQ_In_Sen_Work_A_Pos_01)), PT := T#5s);
Ins_A_Cv_M[6] := Ins_A_Cv_T[1].Q;
Out_CYS_Pos_01_Stopper_A_F_Auto[1] := _p9 AND NOT TimerQ_In_Sen_Work_A_Pos_01;

